(* IEC 61131-3 sources: beedance/reference (part 3) *)

FUNCTION CAUCHY : REAL
VAR_INPUT
	X : REAL;
	T : REAL;
	U : REAL;
END_VAR
VAR
	tmp: REAL;
END_VAR

tmp := x - t;
CAUCHY := math.PI_INV * U / (U*U + tmp*tmp);

(* revision hisdtory
hm	26. oct. 2008	rev 1.0
	original version

*)
END_FUNCTION

FUNCTION CAUCHYCD : REAL
VAR_INPUT
	X : REAL;
	T : REAL;
	U : REAL;
END_VAR

CAUCHYCD := 0.5 + math.PI_INV * ATAN((X - T) / U);

(* revision hisdtory
hm	26. oct. 2008	rev 1.0
	original version

*)
END_FUNCTION

FUNCTION CEIL : INT
VAR_INPUT
	X : REAL;
END_VAR

CEIL := REAL_TO_INT(x);
IF CEIL < X THEN
	CEIL := CEIL + 1;
END_IF;

END_FUNCTION

FUNCTION CEIL2 : DINT
VAR_INPUT
	X : REAL;
END_VAR

CEIL2 := REAL_TO_DINT(X);
IF DINT_TO_REAL(CEIL2) < X THEN
	CEIL2 := CEIL2 + 1;
END_IF;

END_FUNCTION

FUNCTION CMP : BOOL
VAR_INPUT
	X,Y : REAL;
	N : INT;
END_VAR
VAR
	tmp : REAL;
END_VAR

tmp := ABS(x);
IF tmp > 0.0 THEN
	tmp := EXP10(INT_TO_REAL(FLOOR(LOG(tmp))-N+1));
ELSE
	tmp := EXP10(tmp);
END_IF;
CMP := ABS(X - Y) < tmp;

END_FUNCTION

FUNCTION COSH : REAL
VAR_INPUT
	X : REAL;
END_VAR
VAR
	t: REAL;
END_VAR

T := EXP(X);
COSH := (1.0 / T + T) * 0.5;

(* revision histroy
hm	12.1.2007	rev 1.0
	original version

hm	1.12.2007	rev 1.1
	changed code to improve performance

hm	5. jan 2008	rev 1.2
	further performance improvement

hm	10. mar. 2009	rev 1.3
	real constants updated to new systax using dot
*)
END_FUNCTION

FUNCTION COTH : REAL
VAR_INPUT
	X : REAL;
END_VAR

IF X > 20.0 THEN
	COTH :=1.0;
ELSIF X < -20.0 THEN
	COTH := -1.0;
ELSE
	COTH := 1.0 + 2.0 / (EXP(X * 2.0) - 1.0);
END_IF;

(* revision histroy
hm		12.1.2007	rev 1.0
	original version

hm	1.12.2007		rev 1.1
	changed code to improve performance

hm	8. jan 2008	rev 1.2
	further improvement in performance

hm	10. mar 2008	rev 1.3
	extended range of valid inputs to +/- INV
	changed formula for better accuracy

hm	10. mar. 2009	rev 1.4
	real constants updated to new systax using dot
*)
END_FUNCTION

FUNCTION D_TRUNC : DINT
VAR_INPUT
	X : REAL;
END_VAR

D_TRUNC := REAL_TO_DINT(X);
IF X > 0.0 THEN
	IF DINT_TO_REAL(D_TRUNC) > X THEN D_TRUNC := D_TRUNC - 1; END_IF;
ELSE
	IF DINT_TO_REAL(D_TRUNC) < X THEN D_TRUNC := D_TRUNC + 1; END_IF;
END_IF;

(* for systems that support a dint truncation this routine can be replaced by trunc() *)
END_FUNCTION

FUNCTION DEC1 : INT
VAR_INPUT
	X : INT;
	N : INT;
END_VAR

IF X = 0 THEN
	DEC1 := N - 1;
ELSE
	DEC1 := X - 1;
END_IF;

(* this is a very elegant version but 50% slower
X := (X - 1 + N) MOD N;
*)
END_FUNCTION

FUNCTION DEG : REAL
VAR_INPUT
	rad : REAL;
END_VAR

DEG := MODR(57.29577951308232 * RAD, 360.0);
END_FUNCTION

FUNCTION DIFFER : BOOL
VAR_INPUT
	in1 : REAL;
	in2 : REAL;
	X : REAL;
END_VAR

DIFFER := ABS(in1 - in2) > X;
END_FUNCTION

FUNCTION ERF : REAL
VAR_INPUT
	X : REAL;
END_VAR
VAR
	x2 : REAL;
	ax2 : REAL;
END_VAR

x2 := X*X;
ax2 := 0.147 * x2 + 1.0;
ERF := SQRT(1.0 - EXP(-X2 * ((0.27323954473516 + aX2)/(ax2)))) * SGN(x);
END_FUNCTION

FUNCTION ERFC : REAL
VAR_INPUT
	X : REAL;
END_VAR

ERFC := 1.0 - ERF(X);
END_FUNCTION

FUNCTION EVEN : BOOL
VAR_INPUT
	in : DINT;
END_VAR

EVEN := NOT in.0;
END_FUNCTION

FUNCTION EXP10 : REAL
VAR_INPUT
	X : REAL;
END_VAR

EXP10 := EXP(X * 2.30258509299405);
END_FUNCTION

FUNCTION EXPN : REAL
VAR_INPUT
	X : REAL;
	N : INT;
END_VAR
VAR
	sign: BOOL;
END_VAR
VAR
	X_work : REAL;
	N_work : INT;
END_VAR
(* IEC 61131-3 does not let a POU assign to its inputs, so the body works on copies. *)
X_work := X;
N_work := N;

sign := N_work.15;
N_work := ABS(N_work);
IF N_work.0 THEN EXPN := X_work; ELSE EXPN := 1.0; END_IF;
N_work := N_work / 2;
WHILE N_work > 0 DO
   X_work := X_work * X_work;
   IF N_work.0 THEN EXPN := EXPN * X_work; END_IF;
   N_work := N_work / 2;
END_WHILE;
IF sign THEN EXPN := 1.0 / EXPN; END_IF;
END_FUNCTION

FUNCTION FACT : DINT
VAR_INPUT
	X : INT;
END_VAR

IF X >= 0 AND X <= 12 THEN
	FACT := math.FACTS[X];
ELSE
	FACT := -1;
END_IF;

(* working code without array
IF X > 12 OR X < 0 THEN
	FACT := -1;
ELSIF X < 7 THEN
	FACT := 1;
	FOR i := 2 TO X DO
		FACT := FACT * i;
	END_FOR;
ELSE
	FACT := 5040;
	FOR i := 8 TO X DO
		FACT := FACT * i;
	END_FOR;
END_IF;
*)
END_FUNCTION

FUNCTION FIB : DINT
VAR_INPUT
	X : INT;
END_VAR
VAR
	t1, t2: DINT;
END_VAR
VAR
	X_work : INT;
END_VAR
(* IEC 61131-3 does not let a POU assign to its inputs, so the body works on copies. *)
X_work := X;

IF X_work < 0 OR X_work > 46 THEN
	FIB := -1;
ELSIF X_work < 2 THEN
	FIB := X_work;
	RETURN;
ELSE
	(* the fibonacci number is the sum of the two suceeding fibonaci numbers *)
	(* we store the numbers alternatively in t1 and t2 depending on pt *)
	t2 := 1;
	WHILE X_work > 3 DO
		X_work := X_work-2;
		t1 := t1 + t2;
		t2 := t1 + t2;
	END_WHILE;
	IF X_work > 2 THEN t1 := t1 + t2; END_IF;
	fib := t1 + t2;
END_IF;

(* alternative code for very big numbers

IF X < 31 THEN
	fib := 0.4472136 * (expn(1.618034,X) - expn(-0.618034,X));
ELSE
	fib := 0.4472133 * expn(1.618034,X);
END_IF;

*)
END_FUNCTION

FUNCTION FLOOR : INT
VAR_INPUT
	X : REAL;
END_VAR

FLOOR := REAL_TO_INT(X);
IF FLOOR > X THEN
	FLOOR := FLOOR - 1;
END_IF;
END_FUNCTION

FUNCTION FLOOR2 : DINT
VAR_INPUT
	X : REAL;
END_VAR

FLOOR2 := REAL_TO_DINT(X);
IF DINT_TO_REAL(FLOOR2) > X THEN
	FLOOR2 := FLOOR2 - 1;
END_IF;
END_FUNCTION

FUNCTION FRACT : REAL
VAR_INPUT
	x : REAL;
END_VAR

IF ABS(x) < 2.0E9 THEN
	FRACT := x - DINT_TO_REAL(D_TRUNC(x));
ELSE
	FRACT := 0.0;
END_IF;
END_FUNCTION

FUNCTION GAMMA : REAL
VAR_INPUT
	X : REAL;
END_VAR

IF x > 0.0 THEN
	GAMMA := SQRT(math.PI2 / X) * EXPT(math.E_INV * (x + 1.0 / (12.0 * x - 0.1 / X)), X);
END_IF;

(* the stirling formula is not very accurate for small values of X
IF X >=0 THEN GAMMA := SQRT(math.PI2 * X) * EXPT(X / math.E, X); END_IF;
*)
END_FUNCTION

FUNCTION GAUSS : REAL
VAR_INPUT
	X : REAL;
	U : REAL;
	SI: REAL;
END_VAR
VAR
	temp: REAL;
	si_inv: REAL;
END_VAR

temp := X - U;
si_inv := 1.0  / si;
GAUSS := EXP(Temp * Temp * si_inv * si_inv * - 0.5) * 0.39894228 * si_inv;

(* revision hisdtory
hm	6. apr. 2008	rev 1.0
	original version

hm	27. oct. 2008	rev 1.1
	optimized performance

hm	10. mar. 2009	rev 1.2
	real constants updated to new systax using dot

*)
END_FUNCTION

FUNCTION GAUSSCD : REAL
VAR_INPUT
	X : REAL;
	U : REAL;
	SI: REAL;
END_VAR

GAUSSCD := (ERF((X - U) / (SI * 1.414213562)) + 1.0) * 0.5;

(* revision hisdtory
hm	6. apr. 2008	rev 1.0
	original version

hm	10. mar. 2009	rev 1.1
	real constants updated to new systax using dot

*)
END_FUNCTION

FUNCTION GCD : INT
VAR_INPUT
	A : DINT;
	B : DINT;
END_VAR
VAR
	t: DINT;
END_VAR
VAR
	A_work : DINT;
	B_work : DINT;
END_VAR
(* IEC 61131-3 does not let a POU assign to its inputs, so the body works on copies. *)
A_work := A;
B_work := B;

IF A_work = 0 THEN
	GCD := DINT_TO_INT(ABS(B_work));
ELSIF B_work = 0 THEN
	GCD := DINT_TO_INT(ABS(A_work));
ELSE
	A_work := ABS(A_work);
	B_work := ABS(B_work);
	GCD := 1;
	WHILE NOT(A_work.0 OR B_work.0) DO
		A_work := A_work / 2;
		B_work := B_work / 2;
		GCD := GCD * 2;
	END_WHILE;
	WHILE A_work > 0 DO
		IF NOT(A_work.0) THEN A_work := A_work / 2;
		ELSIF NOT(B_work.0) THEN B_work := B_work / 2;
		ELSE
			t:= ABS(A_work-B_work) / 2;
			IF A_work < B_work THEN B_work := t; ELSE A_work := T; END_IF;
		END_IF;
	END_WHILE;
	GCD := GCD * DINT_TO_INT(B_work);
END_IF;
END_FUNCTION

FUNCTION GDF : REAL
VAR_INPUT
	X : REAL;
END_VAR

IF X = 0.0 THEN
	GDF := 0.0;
ELSIF X > 15.0 THEN
	GDF := math.PI05;
ELSIF X < -15.0 THEN
	GDF := -math.PI05;
ELSE
	GDF := ATAN(EXP(X)) * 2.0 - math.PI05;
END_IF;

END_FUNCTION

FUNCTION GOLD : REAL
VAR_INPUT
	X : REAL;
END_VAR

GOLD := (X + SQRT(X*X + 4.0)) * 0.5;

END_FUNCTION

FUNCTION HYPOT : REAL
VAR_INPUT
	X : REAL;
	Y : REAL;
END_VAR

HYPOT := SQRT(x*x + y*y);

END_FUNCTION

FUNCTION INC : INT
VAR_INPUT
	X : INT;
	D : INT;
	M : INT;
END_VAR

INC := (X + D + M + 1) MOD (M + 1);
END_FUNCTION

FUNCTION INC1 : INT
VAR_INPUT
	X : INT;
	N : INT;
END_VAR

IF X >= N - 1 THEN
	INC1 := 0;
ELSE
	INC1 := X + 1;
END_IF;
END_FUNCTION

FUNCTION INC2 : INT
VAR_INPUT
	X : INT;
	D : INT;
	L : INT;
	U : INT;
END_VAR
VAR
	tmp: INT;
END_VAR

tmp := U - L + 1;
INC2 := (X + D - L + tmp) MOD tmp + L;
END_FUNCTION

FUNCTION INV : REAL
VAR_INPUT
	X : REAL;
END_VAR

IF X <> 0.0 THEN INV := 1.0 / X; END_IF;

END_FUNCTION

// Commented out for beedance: it uses REAL_TO_DW, which is commented out.
// FUNCTION LAMBERT_W : REAL
// VAR_INPUT
// 	X : REAL;
// END_VAR
// VAR
// 	w : REAL;
// 	i : INT;
// 	we: REAL;
// 	w1e: REAL;
// 	last: DWORD;
// 	ewx: REAL;
// END_VAR
//
// (* check for valid input and return -1000 if too low *)
// IF x < -0.367879441171442 THEN
// 	LAMBERT_W := -1000.0;
// 	RETURN;
// (* return 0 if x = 0 *)
// ELSIF x = 0.0 THEN
// 	RETURN;
// (* first an estimate is calculated *)
// ELSIF x <= 500.0 THEN
// 	w := LN(x + 1.0);
// 	w := 0.665 * (1.0 + 0.0195 * w) * w + 0.04;
// ELSE
// 	w := LN(x - 4.0) - (1.0 - 1.0/LN(x)) * LN(LN(x));
// END_IF;
// (* use estimate to calculate exact result *)
// FOR i := 0 TO 5 DO
// 	ewx := EXP(w);
// 	we := w * ewx - x;
// 	w1e := (w+1.0) * ewx;
// 	last := REAL_TO_DW(w) AND 16#FFFF_FFFC;
// 	w := w - (we / (w1e - (w+2.0) * we / (2.0 * w + 2.0)));
// 	IF (REAL_TO_DW(w) AND 16#FFFF_FFFC) = last THEN EXIT; END_IF;
// END_FOR;
// LAMBERT_W := w;
//
//
// (* revision hisdtory
// hm	26. oct. 2008	rev 1.0
// 	original version
//
// hm	10. mar. 2009	rev 1.1
// 	real constants updated to new systax using dot
//
// *)
// END_FUNCTION

FUNCTION LANGEVIN : REAL
VAR_INPUT
	X : REAL;
END_VAR

IF X = 0.0 THEN
	LANGEVIN := 0.0;
ELSE
	LANGEVIN := COTH(X) - 1.0 / X;
END_IF;
END_FUNCTION

FUNCTION MAX3 : REAL
VAR_INPUT
	in1 : REAL;
	in2 : REAL;
	in3 : REAL;
END_VAR

MAX3 := MAX(MAX(IN1,IN2),IN3);
END_FUNCTION

FUNCTION MID3 : REAL
VAR_INPUT
	IN1 : REAL;
	IN2 : REAL;
	IN3 : REAL;
END_VAR
VAR
	IN1_work : REAL;
	IN2_work : REAL;
END_VAR
(* IEC 61131-3 does not let a POU assign to its inputs, so the body works on copies. *)
IN1_work := IN1;
IN2_work := IN2;

IF IN1_work > IN2_work THEN MID3 := IN1_work; IN1_work := IN2_work; IN2_work := MID3; END_IF;
IF IN2_work > IN3 THEN IN2_work := IN3; END_IF;
MID3 := SEL(IN1_work > IN2_work, IN2_work, IN1_work);

(*
hm	1.1.2007	rev 1.1
	rewrote the function for better performance

hm	18. mar. 2011	rev 1.2
	improve performance
*)
END_FUNCTION

FUNCTION MIN3 : REAL
VAR_INPUT
	in1 : REAL;
	in2 : REAL;
	in3 : REAL;
END_VAR

MIN3 := MIN(MIN(IN1,IN2),IN3);
END_FUNCTION

FUNCTION MODR : REAL
VAR_INPUT
	IN : REAL;
	DIVI : REAL;
END_VAR

IF divi = 0.0 THEN
	MODR := 0.0;
ELSE
	MODR := in - DINT_TO_REAL(FLOOR2(in / divi)) * divi;
END_IF;
END_FUNCTION

FUNCTION MUL_ADD : REAL
VAR_INPUT
	X : REAL;
	K : REAL;
	O : REAL;
END_VAR

MUL_ADD := X * K + O;
END_FUNCTION

FUNCTION NEGX : REAL
VAR_INPUT
	X : REAL;
END_VAR

NEGX := -X;

END_FUNCTION

FUNCTION RAD : REAL
VAR_INPUT
	DEG : REAL;
END_VAR

RAD := MODR(0.0174532925199433 * DEG, math.PI2);
END_FUNCTION

FUNCTION RDM : REAL
VAR_INPUT
	last : REAL;
END_VAR
VAR
	tn : DWORD;
	tc : INT;
END_VAR

tn := T_PLC_MS();
tc := BIT_COUNT(tn);
tn.31 := tn.2;
tn.30 := tn.5;
tn.29 := tn.4;
tn.28 := tn.1;
tn.27 := tn.0;
tn.26 := tn.7;
tn.25 := tn.6;
tn.24 := tn.3;
tn := ROL(tn,BIT_COUNT(tn)) OR 16#80000001;
tn := ULINT_TO_DWORD(DWORD_TO_ULINT(tn) MOD 71474513 + INT_TO_ULINT(tc + 77));
RDM := FRACT(DWORD_TO_REAL(tn) / 10000000.0 * (math.E - LIMIT(0.0,last,1.0)));

(*
pt := ADR(temp);
pt^ := (T_PLC_MS() AND 16#007FFFFF) OR 16#3D000000;
RDM := fract(modR(temp*e+pi1, PI1-last) + modR(temp*PI1+e + last,e-last));
*)
END_FUNCTION

FUNCTION RDM2 : INT
VAR_INPUT
	last : INT;
	low : INT;
	high : INT;
END_VAR

RDM2 := TRUNC(RDM(FRACT(last * math.PI)) * (high - low + 1)) + low;
END_FUNCTION

FUNCTION RDMDW : DWORD
VAR_INPUT
	last : DWORD;
END_VAR
VAR
	RX: REAL;
	M: REAL;
END_VAR

M := BIT_COUNT(last);
RX := RDM(FRACT(M * math.PI));
RDMDW := SHL(REAL_TO_DWORD(rx*65535),16);
RX := RDM(FRACT(M * math.E));
RDMDW := RDMDW OR (REAL_TO_DWORD(rx*65535) AND 16#0000FFFF);
END_FUNCTION

FUNCTION REAL_TO_FRAC : FRACTION
VAR_INPUT
	X : REAL;					(* in einen Bruch umzuwandelnder Wert *)
	N : INT;					(* maximale Größe des Nenners *)
END_VAR
VAR
	temp : DINT;				(* Merker für Berechnungen *)

	sign: BOOL;					(* Vorzeichen vom Eingangswert *)
	X_gerundet: DINT;			(* Wert von Bruch, auf ganze Zahl gerundet *)
	X_ohne_Nachkomma: REAL;		(* Wert von Bruch, ohne Nachkommastellen *)
	Numerator:       DINT := 1;	(* Initialwert Zaehler  *)
	Denominator:     DINT := 0;	(* Initialwert Nenner *)
	Numerator_old:   DINT := 0;	(* Initialwert Zaehler der letzten Berechnung  *)
	Denominator_old: DINT := 1;	(* Initialwert Zaehler der letzten Berechnung   *)

END_VAR
VAR
	X_work : REAL;
END_VAR
(* IEC 61131-3 does not let a POU assign to its inputs, so the body works on copies. *)
X_work := X;

IF X_work < 0.0 THEN
	sign := TRUE;								(* Vorzeichen merken *)
	X_work := ABS(X_work);								(* Absolutwert berechnen *)
END_IF;

REPEAT
	X_gerundet := REAL_TO_DINT(X_work);

	(* Zaehler berechnen *)
	temp := numerator * X_gerundet + numerator_old;		(* Zaehler um Vorkammawert erweitern *)
	numerator_old := numerator;							(* Zaehler der letzten Berechnung speichern *)
	numerator := temp;									(* Zaehler dieser Berechnung speichern *)

	(* Nenner berechnen *)
	temp := denominator * X_gerundet + denominator_old;	(* Nenner um Vorkammawert erweitern *)
	denominator_old := denominator;						(* Nenner der letzten Berechnung speichern *)
	denominator := temp;								(* Nenner dieser Berechnung speichern *)

	(* Restwert berechnen *)
	X_ohne_Nachkomma := DINT_TO_REAL(X_gerundet);
	IF X_work = X_ohne_Nachkomma THEN						(* Bruch geht ohne Rest auf *)
		IF ABS(denominator) <= N THEN						(* kein Rundungsfehler *)
			numerator_old := numerator;					(* Numerator_old wird von Funktion zurückgegeben *)
			denominator_old := denominator;			(* Denominator_old wird von Funktion zurückgegeben *)
		END_IF
		EXIT;											(* keine weitere Berechnung notwendig *)
	ELSE
		X_work := 1.0 / (X_work - X_ohne_Nachkomma);				(* Kehrwert vom Rest -> Neuer Bruch *)
	END_IF

UNTIL
	ABS(Denominator) > N
END_REPEAT

(* correct sign if X was negative *)
IF sign THEN
	REAL_TO_FRAC.NUMERATOR := -1 * ABS(DINT_TO_INT(numerator_old));
ELSE
	REAL_TO_FRAC.NUMERATOR :=  ABS(DINT_TO_INT(numerator_old));
END_IF
REAL_TO_FRAC.DENOMINATOR := ABS(DINT_TO_INT(denominator_old));
END_FUNCTION

FUNCTION RND : REAL
VAR_INPUT
	X : REAL;
	N : INT;
END_VAR
VAR
	M : REAL;
END_VAR

IF X = 0.0 THEN
	RND := 0.0;
ELSE
	M := EXPN(10.0,N - CEIL(LOG(ABS(X))));
	RND := DINT_TO_REAL(REAL_TO_DINT(X * M)) / M;
END_IF;

END_FUNCTION

 FUNCTION ROUND : REAL
VAR_INPUT
	in : REAL;
	N : INT;
END_VAR
VAR
	X: REAL;
END_VAR

X := setup.DECADES[LIMIT(0,N,8)];
ROUND := DINT_TO_REAL(REAL_TO_DINT(in * X)) / X;

END_FUNCTION

FUNCTION SGN : INT
VAR_INPUT
	X : REAL;
END_VAR

IF X > 0 THEN
	SGN := 1;
ELSIF X < 0 THEN
	SGN := -1;
ELSE
	SGN := 0;
END_IF;

(* revision histroy
hm	16. oct 2007	rev 1.0
	original version

hm	11. nov 2007	rev 1.1
	changed type of function from real to int

*)
END_FUNCTION

FUNCTION SIGMOID : REAL
VAR_INPUT
	X : REAL;
END_VAR

IF X > 20.0 THEN
	SIGMOID := 1.0;
ELSIF x < -85.0 THEN
	SIGMOID := 0.0;
ELSE
	SIGMOID := 1.0 / (1.0 + EXP(-X));
END_IF;
END_FUNCTION

FUNCTION SIGN_I : BOOL
VAR_INPUT
	IN : DINT;
END_VAR

SIGN_I := in.31;
END_FUNCTION

FUNCTION SIGN_R : BOOL
VAR_INPUT
	in : REAL;
END_VAR

SIGN_R := in < 0.0;
END_FUNCTION

FUNCTION SINC : REAL
VAR_INPUT
	X : REAL;
END_VAR

IF X = 0.0 THEN
	SINC := 1.0;
ELSE
	SINC := SIN(x) / x;
END_IF;

(* revision histroy
hm	11. mar. 2008	rev 1.0
	original version

hm	1.12.2007	rev 1.1
	changed code to improove performance

hm 10. mar. 2009	rev 1.2
	real constants updated to new systax using dot

*)
END_FUNCTION

FUNCTION SINH : REAL
VAR_INPUT
	X : REAL;
END_VAR

IF ABS(x) < 2E-3 THEN
	SINH := X;
ELSE
	SINH := (EXP(x) - EXP(-x)) * 0.5;
END_IF;
END_FUNCTION

FUNCTION SQRTN : REAL
VAR_INPUT
	X : REAL;
	N : INT;
END_VAR

IF N > 0 THEN
	SQRTN := EXP(LN(x) / INT_TO_REAL(n));
ELSE
	SQRTN := 0.0;
END_IF;
END_FUNCTION

FUNCTION TANC : REAL
VAR_INPUT
	X : REAL;
END_VAR

IF X = 0.0 THEN
	TANC := 1.0;
ELSE
	TANC := TAN(x) / x;
END_IF;

(* revision histroy
hm	23. oct. 2008	rev 1.0
	original version

hm 10. mar. 2009	rev 1.1
	real constants updated to new systax using dot

*)
END_FUNCTION

FUNCTION TANH : REAL
VAR_INPUT
	X : REAL;
END_VAR

IF X > 20.0 THEN
	TANH := 1.0;
ELSIF X < -20.0 THEN
	TANH := -1.0;
ELSE
	TANH := 1.0 - 2.0 / (EXP(2.0 * x) + 1.0);
END_IF;

(* revision hisdtory
hm		12.1.2007		rev 1.0
	original version

hm		1.12.2007		rev 1.1
	changed code to improve performance

hm		10. mar 2008	rev 1.2
	corrected an error in formula
	extended range of valid inputs to +/- INV

hm 10. mar. 2009	rev 1.3
	real constants updated to new systax using dot

*)
END_FUNCTION

FUNCTION WINDOW : BOOL
VAR_INPUT
	low : REAL;
	in : REAL;
	high : REAL;
END_VAR

WINDOW := in < high AND in > low;
END_FUNCTION

FUNCTION WINDOW2 : BOOL
VAR_INPUT
	LOW : REAL;
	IN : REAL;
	HIGH : REAL;
END_VAR

WINDOW2 := IN >= LOW AND IN <= HIGH;
END_FUNCTION

FUNCTION_BLOCK ESR_COLLECT
VAR_INPUT
	ESR_0, ESR_1, ESR_2, ESR_3, ESR_4, ESR_5, ESR_6, ESR_7 : ARRAY [0..3] OF esr_data;
	rst : BOOL;
END_VAR
VAR_IN_OUT
	pos : INT;
END_VAR
VAR_OUTPUT
	ESR_OUT : ARRAY[0..31] OF esr_data;
END_VAR
VAR CONSTANT
	max_in : INT := 3; (* max limit of input array *)
	max_out : INT := 32; (* number of elements in array *)
END_VAR
VAR
	cnt : INT := -1;
END_VAR

IF rst OR cnt < 0 THEN
	pos := -1;
ELSE
	FOR cnt := 0 TO max_in DO
	IF esr_0[cnt].typ > 0 THEN pos := INC1(pos, max_out); esr_out[pos] := esr_0[cnt]; END_IF;
	IF esr_1[cnt].typ > 0 THEN pos := INC1(pos, max_out); esr_out[pos] := esr_1[cnt]; END_IF;
	IF esr_2[cnt].typ > 0 THEN pos := INC1(pos, max_out); esr_out[pos] := esr_2[cnt]; END_IF;
	IF esr_3[cnt].typ > 0 THEN pos := INC1(pos, max_out); esr_out[pos] := esr_3[cnt]; END_IF;
	IF esr_4[cnt].typ > 0 THEN pos := INC1(pos, max_out); esr_out[pos] := esr_4[cnt]; END_IF;
	IF esr_5[cnt].typ > 0 THEN pos := INC1(pos, max_out); esr_out[pos] := esr_5[cnt]; END_IF;
	IF esr_6[cnt].typ > 0 THEN pos := INC1(pos, max_out); esr_out[pos] := esr_6[cnt]; END_IF;
	IF esr_7[cnt].typ > 0 THEN pos := INC1(pos, max_out); esr_out[pos] := esr_7[cnt]; END_IF;
   END_FOR;
END_IF;
END_FUNCTION_BLOCK

FUNCTION_BLOCK ESR_MON_B8
VAR_INPUT
	s0, s1, s2, s3, s4, s5, s6, s7 : BOOL;
	DT_in : DT;
END_VAR
VAR_INPUT CONSTANT
	a0, a1, a2, a3, a4, a5, a6, a7 : STRING(10);
END_VAR
VAR_OUTPUT
	ESR_Flag : BOOL;
END_VAR
VAR_IN_OUT
	ESR_Out: ARRAY [0..3] OF esr_data;
END_VAR
VAR
	x0, x1, x2, x3, x4, x5, x6, x7 : BOOL;
	tx: TIME;
	cnt : INT;
END_VAR

(* read system timer *)
tx := DWORD_TO_TIME(T_PLC_MS());

ESR_Flag := FALSE;
esr_out[3].typ := 0;
esr_out[2].typ := 0;
esr_out[1].typ := 0;
esr_out[0].typ := 0;
cnt := 0;

(* check if inputs have chaged and fill buffer *)
IF s0 <> X0 THEN
	esr_out[cnt].typ := USINT_TO_BYTE(10 + BOOL_TO_USINT(s0));
	esr_out[cnt].adress := a0;
	esr_out[cnt].DS := DT_in;
	esr_out[cnt].TS := TX;
	X0 := S0;
	cnt := cnt + 1;
	esr_flag := TRUE;
END_IF;
IF s1 <> X1 THEN
	esr_out[cnt].typ := USINT_TO_BYTE(10 + BOOL_TO_USINT(s1));
	esr_out[cnt].adress := a1;
	esr_out[cnt].DS := DT_in;
	esr_out[cnt].TS := TX;
	X1 := S1;
	cnt := cnt + 1;
	esr_flag := TRUE;
END_IF;
IF s2 <> X2 THEN
	esr_out[cnt].typ := USINT_TO_BYTE(10 + BOOL_TO_USINT(s2));
	esr_out[cnt].adress := a2;
	esr_out[cnt].DS := DT_in;
	esr_out[cnt].TS := TX;
	X2 := S2;
	cnt := cnt + 1;
	esr_flag := TRUE;
END_IF;
IF s3 <> X3 THEN
	esr_out[cnt].typ := USINT_TO_BYTE(10 + BOOL_TO_USINT(s3));
	esr_out[cnt].adress := a3;
	esr_out[cnt].DS := DT_in;
	esr_out[cnt].TS := TX;
	X3 := S3;
	cnt := cnt + 1;
	esr_flag := TRUE;
END_IF;
IF s4 <> X4 AND cnt < 4 THEN
	esr_out[cnt].typ := USINT_TO_BYTE(10 + BOOL_TO_USINT(s4));
	esr_out[cnt].adress := a4;
	esr_out[cnt].DS := DT_in;
	esr_out[cnt].TS := TX;
	X4 := S4;
	cnt := cnt + 1;
	esr_flag := TRUE;
END_IF;
IF s5 <> X5  AND cnt < 4 THEN
	esr_out[cnt].typ := USINT_TO_BYTE(10 + BOOL_TO_USINT(s5));
	esr_out[cnt].adress := a5;
	esr_out[cnt].DS := DT_in;
	esr_out[cnt].TS := TX;
	X5 := S5;
	cnt := cnt + 1;
	esr_flag := TRUE;
END_IF;
IF s6 <> X6  AND cnt < 4 THEN
	esr_out[cnt].typ := USINT_TO_BYTE(10 + BOOL_TO_USINT(s6));
	esr_out[cnt].adress := a6;
	esr_out[cnt].DS := DT_in;
	esr_out[cnt].TS := TX;
	X6 := S6;
	cnt := cnt + 1;
	esr_flag := TRUE;
END_IF;
IF s7 <> X7  AND cnt < 4 THEN
	esr_out[cnt].typ := USINT_TO_BYTE(10 + BOOL_TO_USINT(s7));
	esr_out[cnt].adress := a7;
	esr_out[cnt].DS := DT_in;
	esr_out[cnt].TS := TX;
	X7 := S7;
	cnt := cnt + 1;
	esr_flag := TRUE;
END_IF;
END_FUNCTION_BLOCK

// Commented out for beedance: it reads the bits of a REAL as a DWORD, or back, through a pointer; a beedance reference (REF_TO) refers to a variable of its own type.
// FUNCTION_BLOCK ESR_MON_R4
// VAR_INPUT
// 	R0, R1, R2, R3 : REAL;
// 	DT_in : DT;
// END_VAR
// VAR_INPUT CONSTANT
// 	a0, a1, a2, a3 : STRING(10);
// 	s0, s1, s2, s3 : REAL;
// END_VAR
// VAR_OUTPUT
// 	ESR_Flag : BOOL;
// END_VAR
// VAR_IN_OUT
// 	ESR_Out: ARRAY [0..3] OF esr_data;
// END_VAR
// VAR
// 	p0, p1, p2, p3 : REF_TO DWORD;
// 	x0, x1, x2, x3 : REAL;
// 	tx: TIME;
// 	cnt : INT;
// END_VAR
//
//
// (* read system timer *)
// tx := DWORD_TO_TIME(T_PLC_MS());
// P0 := REF(R0);
// P1 := REF(R1);
// P2 := REF(R2);
// P3 := REF(R3);
//
// ESR_Flag := FALSE;
// esr_out[3].typ := 0;
// esr_out[2].typ := 0;
// esr_out[1].typ := 0;
// esr_out[0].typ := 0;
// cnt := 0;
//
// (* check if inputs have chaged and fill buffer *)
// IF DIFFER(R0,  X0, S0) THEN
// 	esr_out[cnt].typ := 20;
// 	esr_out[cnt].adress := a0;
// 	esr_out[cnt].DS := DT_in;
// 	esr_out[cnt].TS := TX;
// 	esr_out[cnt].data[0] := Byte_of_Dword(P0^,0);
// 	esr_out[cnt].data[1] := Byte_of_Dword(P0^,1);
// 	esr_out[cnt].data[2] := Byte_of_Dword(P0^,2);
// 	esr_out[cnt].data[3] := Byte_of_Dword(P0^,3);
// 	X0 := R0;
// 	cnt := cnt + 1;
// 	esr_flag := TRUE;
// END_IF;
// IF differ(R1,  X1, S1) THEN
// 	esr_out[cnt].typ := 20;
// 	esr_out[cnt].adress := a1;
// 	esr_out[cnt].DS := DT_in;
// 	esr_out[cnt].TS := TX;
// 	esr_out[cnt].data[0] := Byte_of_Dword(P1^,0);
// 	esr_out[cnt].data[1] := Byte_of_Dword(P1^,1);
// 	esr_out[cnt].data[2] := Byte_of_Dword(P1^,2);
// 	esr_out[cnt].data[3] := Byte_of_Dword(P1^,3);
// 	X1 := R1;
// 	cnt := cnt + 1;
// 	esr_flag := TRUE;
// END_IF;
// IF differ(R2,  X2, S2) THEN
// 	esr_out[cnt].typ := 20;
// 	esr_out[cnt].adress := a2;
// 	esr_out[cnt].DS := DT_in;
// 	esr_out[cnt].TS := TX;
// 	esr_out[cnt].data[0] := Byte_of_Dword(P2^,0);
// 	esr_out[cnt].data[1] := Byte_of_Dword(P2^,1);
// 	esr_out[cnt].data[2] := Byte_of_Dword(P2^,2);
// 	esr_out[cnt].data[3] := Byte_of_Dword(P2^,3);
// 	X2 := R2;
// 	cnt := cnt + 1;
// 	esr_flag := TRUE;
// END_IF;
// IF DIFFER(R3,  X3, S3) THEN
// 	esr_out[cnt].typ := 20;
// 	esr_out[cnt].adress := a3;
// 	esr_out[cnt].DS := DT_in;
// 	esr_out[cnt].TS := TX;
// 	esr_out[cnt].data[0] := Byte_of_Dword(P3^,0);
// 	esr_out[cnt].data[1] := Byte_of_Dword(P3^,1);
// 	esr_out[cnt].data[2] := Byte_of_Dword(P3^,2);
// 	esr_out[cnt].data[3] := Byte_of_Dword(P3^,3);
// 	X3 := R3;
// 	cnt := cnt + 1;
// 	esr_flag := TRUE;
// END_IF;
//
// END_FUNCTION_BLOCK

FUNCTION_BLOCK ESR_MON_X8
VAR_INPUT
	s0, s1, s2, s3, s4, s5, s6, s7 : BYTE;
	DT_in : DT;
	Mode : BYTE := 3;
END_VAR
VAR_INPUT CONSTANT
	a0, a1, a2, a3, a4, a5, a6, a7 : STRING(10);
END_VAR
VAR_OUTPUT
	ESR_Flag : BOOL;
END_VAR
VAR_IN_OUT
	ESR_Out: ARRAY [0..3] OF esr_data;
END_VAR
VAR
	x0, x1, x2, x3, x4, x5, x6, x7 : BYTE;
	tx: TIME;
	cnt : INT;
END_VAR

(* read system timer *)
tx := DWORD_TO_TIME(T_PLC_MS());

ESR_Flag := FALSE;
esr_out[3].typ := 0;
esr_out[2].typ := 0;
esr_out[1].typ := 0;
esr_out[0].typ := 0;
cnt := 0;

(* check if inputs have chaged and fill buffer *)
IF s0 <> X0 AND ((s0 < 100) OR (S0 > 99 AND S0 < 200 AND mode >= 2) OR (S0 > 199 AND mode = 3)) THEN
	esr_out[cnt] := status_to_ESR(s0, a0, DT_in, TX);
	X0 := S0;
	cnt := cnt + 1;
	esr_flag := TRUE;
END_IF;
IF s1 <> X1 AND ((s1 < 100) OR (S1 > 99 AND S1 < 200 AND mode >= 2) OR (S1 > 199 AND mode = 3)) THEN
	esr_out[cnt] := status_to_ESR(s1, a1, DT_in, TX);
	X1 := S1;
	cnt := cnt + 1;
	esr_flag := TRUE;
END_IF;
IF s2 <> X2 AND ((s2 < 100) OR (S2 > 99 AND S2 < 200 AND mode >= 2) OR (S2 > 199 AND mode = 3)) THEN
	esr_out[cnt] := status_to_ESR(s2, a2, DT_in, TX);
	X2 := S2;
	cnt := cnt + 1;
	esr_flag := TRUE;
END_IF;
IF s3 <> X3 AND ((s3 < 100) OR (S3 > 99 AND S3 < 200 AND mode >= 2) OR (S3 > 199 AND mode = 3)) THEN
	esr_out[cnt] := status_to_ESR(s3, a3, DT_in, TX);
	X3 := S3;
	cnt := cnt + 1;
	esr_flag := TRUE;
END_IF;
IF cnt < 4 AND s4 <> X4 AND ((s4 < 100) OR (S4 > 99 AND S4 < 200 AND mode >= 2) OR (S4 > 199 AND mode = 3)) THEN
	esr_out[cnt] := status_to_ESR(s4, a4, DT_in, TX);
	X4 := S4;
	cnt := cnt + 1;
	esr_flag := TRUE;
END_IF;
IF cnt < 4 AND s5 <> X5 AND ((s5 < 100) OR (S5 > 99 AND S5 < 200 AND mode >= 2) OR (S5 > 199 AND mode = 3)) THEN
	esr_out[cnt] := status_to_ESR(s5, a5, DT_in, TX);
	X5 := S5;
	cnt := cnt + 1;
	esr_flag := TRUE;
END_IF;
IF cnt < 4 AND s6 <> X6 AND ((s6 < 100) OR (S6 > 99 AND S6 < 200 AND mode >= 2) OR (S6 > 199 AND mode = 3)) THEN
	esr_out[cnt] := status_to_ESR(s6, a6, DT_in, TX);
	X6 := S6;
	cnt := cnt + 1;
	esr_flag := TRUE;
END_IF;
IF cnt < 4 AND s7 <> X7 AND ((s7 < 100) OR (S7 > 99 AND S7 < 200 AND mode >= 2) OR (S7 > 199 AND mode = 3)) THEN
	esr_out[cnt] := status_to_ESR(s7, a7, DT_in, TX);
	X7 := S7;
	cnt := cnt + 1;
	esr_flag := TRUE;
END_IF;
END_FUNCTION_BLOCK

FUNCTION OSCAT_VERSION : DWORD
VAR_INPUT
	IN : BOOL;
END_VAR

IF in THEN
	OSCAT_VERSION := DATE_TO_DWORD(D#2024-07-16);
ELSE
	OSCAT_VERSION := 335;
END_IF;
END_FUNCTION

FUNCTION STATUS_TO_ESR : esr_data
VAR_INPUT
	status : BYTE;
	adress : STRING(10);
	DT_in : DT;
	TS : TIME;
END_VAR

IF status < 100 THEN
	status_to_ESR.typ := 1;
ELSIF status < 200 THEN
	status_to_ESR.typ := 2;
ELSE
	status_to_ESR.typ := 3;
END_IF;
status_to_ESR.adress:= adress;
status_to_ESR.DS := DT_in;
status_to_ESR.TS := TS;
status_to_ESR.data[0] := status;

END_FUNCTION

// Commented out for beedance: it reads or writes the bytes of a STRING through a pointer; a beedance reference (REF_TO) refers to a whole variable of its type.
// FUNCTION BIN_TO_BYTE : BYTE
// VAR_INPUT
// 	BIN : STRING(12);
// END_VAR
// VAR
// 	pt : REF_TO BYTE;
// 	i: INT;
// 	X: BYTE;
// 	stop: INT;
// END_VAR
//
// pt := REF(bin);
// stop := LEN(bin);
// FOR I := 1 TO stop DO
// 	x := pt^;
// 	(* calculate the value of the digit *)
// 	IF X = 48 THEN
// 		BIN_TO_BYTE := SHL(BIN_TO_BYTE,1);
// 	ELSIF X = 49 THEN
// 		BIN_TO_BYTE := SHL(BIN_TO_BYTE,1) OR 1;
// 	END_IF;
// 	pt := pt + 1;
// END_FOR;
//
//
//
// (* revision histroy
// hm	18. jun. 2008	rev 1.0
// 	original release
//
// hm	20. sep. 2008	rev 1.1
// 	changed length of input string from 20 to 12
//
// hm	26. jul. 2009	rev 1.2
// 	optimized code
// *)
//
// END_FUNCTION

// Commented out for beedance: it reads or writes the bytes of a STRING through a pointer; a beedance reference (REF_TO) refers to a whole variable of its type.
// FUNCTION BIN_TO_DWORD : DWORD
// VAR_INPUT
// 	BIN : STRING(40);
// END_VAR
// VAR
// 	pt : REF_TO BYTE;
// 	i: INT;
// 	X: BYTE;
// 	stop: INT;
// END_VAR
//
// pt := REF(bin);
// stop := LEN(bin);
// FOR I := 1 TO stop DO
// 	x := pt^;
// 	(* calculate the value of the digit *)
// 	IF X = 48 THEN
// 		BIN_TO_DWORD := SHL(BIN_TO_DWORD,1);
// 	ELSIF X = 49 THEN
// 		BIN_TO_DWORD := SHL(BIN_TO_DWORD,1) OR 1;
// 	END_IF;
// 	pt := pt + 1;
// END_FOR;
//
//
//
// (* revision histroy
// hm	18. jun. 2008	rev 1.0
// 	original release
//
// hm	20. sep. 2008	rev 1.1
// 	changed length of input dtring from 20 to 40
//
// hm	26. jul 2009	rev 1.2
// 	optimized code
// *)
//
// END_FUNCTION

// Commented out for beedance: it reads or writes the bytes of a STRING through a pointer; a beedance reference (REF_TO) refers to a whole variable of its type.
// FUNCTION BYTE_TO_STRB : STRING(8)
// VAR_INPUT
// 	IN : BYTE;
// END_VAR
// VAR
// 	i: INT;
// 	pt : REF_TO BYTE;
// END_VAR
//
//
// (* pointer für die ausgabe ermitteln *)
// pt := REF(BYTE_TO_STRB);
// (* die 8 ausgabecharacter ermitteln und schreiben *)
// FOR i := 1 TO 8 DO
// 	pt^ := BOOL_TO_BYTE(in.7) + 48;
// 	in := SHL(in,1);
// 	pt := pt + 1;
// END_FOR;
//
// (* der ausgabestring muss noch mit 0 abgeschlossen werden *)
// pt^ := 0;
//
// (* code before rev 1.1
// FOR i := 1 TO 8 DO
// 	IF in.0 = 0 THEN temp := CONCAT('0', temp); ELSE temp := CONCAT('1', temp); END_IF;
// 	in := SHR(in, 1);
// END_FOR;
// BYTE_TO_STRB := temp;
// *)
// END_FUNCTION

// Commented out for beedance: it reads or writes the bytes of a STRING through a pointer; a beedance reference (REF_TO) refers to a whole variable of its type.
// FUNCTION BYTE_TO_STRH : STRING(2)
// VAR_INPUT
// 	IN : BYTE;
// END_VAR
// VAR
// 	temp : BYTE;
// 	PT : REF_TO BYTE;
// END_VAR
//
//
// (* read pointer to output string *)
// PT := REF(BYTE_TO_STRH);
// (* calculate high order hex value *)
// temp := SHR(in,4);
// (* convert value to hex character *)
// IF temp <= 9 THEN temp := temp + 48; ELSE temp := temp + 55; END_IF;
// (* write friat character to output string *)
// PT^ := temp;
// (* calculate low order hex value *)
// temp := in AND 2#00001111;
// IF temp <= 9 THEN temp := temp + 48; ELSE temp := temp + 55; END_IF;
// (* increment pointer and wirte low order character *)
// pt := pt + 1;
// pt^ := temp;
// (* set pointer at the end of the output string and close the string with 0 *)
// pt := pt + 1;
// pt^:= 0;
//
//
// (* code before rev 1.2
// FOR i := 1 TO 2 DO
// 	X := in AND 2#1111;
// 	IF X <= 9 THEN X := X + 48; ELSE X := X + 55; END_IF;
// 	Cx := CHR(X);
// 	temp := CONCAT(Cx, temp);
// 	in := SHR(in,4);
// END_FOR;
// BYTE_TO_STRH := temp;
// *)
// END_FUNCTION

// Commented out for beedance: it computes with pointers as addresses (pt := pt + 1); beedance references (REF_TO) have no arithmetic.
// FUNCTION CAPITALIZE : STRING(STRING_LENGTH)
// VAR_INPUT
// 	str : STRING(STRING_LENGTH);
// END_VAR
// VAR
// 	PT : REF_TO BYTE;
// 	pos : INT;
// 	L : INT;
// 	first : BOOL := TRUE;
// END_VAR
//
// PT := REF(CAPITALIZE);
// CAPITALIZE := str;
// L := LEN(str);
// FOR pos := 1 TO l DO
// 	IF first THEN pt^ := TO_UPPER(pt^);	END_IF;
// 	(* remember in first if the next char needs to capitalized *)
// 	first := pt^= 32;
// 	PT := pt + 1;
// END_FOR;
//
// (* revision histroy
// hm		4. mar 2008	rev 1.0
// 	original release
//
// hm	29. mar. 2008	rev 1.1
// 	changed STRING to STRING(STRING_LENGTH)
//
// hm	20. jun. 2008	rev 1.2
// 	improved performance
//
// *)
//
// END_FUNCTION

// Commented out for beedance: it uses CODE, which is commented out.
// FUNCTION CHARCODE : BYTE
// VAR_INPUT
// 	STR : STRING(10);
// END_VAR
// VAR
// 	found: STRING(1);
// 	search : STRING(10);
// 	pos: INT;
// 	i: INT;
// END_VAR
//
// IF LEN(str) = 1 THEN
// 	CHARCODE := CODE(STR, 1);
// ELSIF str <> '' THEN
// 	(* construct search string *)
// 	search := CONCAT('&', str);
// 	search := CONCAT(search, ';');
// 	WHILE pos = 0 AND (i < 4) DO
// 		i := i + 1;
// 		pos := FIND(setup.CHARNAMES[i], search);
// 	END_WHILE;
// 	found := MID(setup.CHARNAMES[i], 1, pos - 1);
// 	CHARCODE := CODE(found, 1);
// END_IF;
//
// END_FUNCTION

// Commented out for beedance: it uses CHR_TO_STRING, which is commented out.
// FUNCTION CHARNAME : STRING(10)
// VAR_INPUT
// 	C : BYTE;
// END_VAR
// VAR
// 	pos: INT;
// 	i : INT;
// END_VAR
//
// IF C <> 0 THEN
// 	(* construct search string from code followed by $ sign, also clear charname string*)
// 	CHARNAME := CHR_TO_STRING(C);
// 	CHARNAME := CONCAT(CHARNAME,'&');
// 	CHARNAME := CONCAT(';', CHARNAME);
// 	WHILE pos = 0 AND (i < 4) DO
// 		i := i + 1;
// 		pos := FIND(setup.CHARNAMES[i], CHARNAME);
// 	END_WHILE;
// 	IF pos > 0 THEN
// 		CHARNAME := MID(setup.CHARNAMES[i], 10, pos + 3);
// 		(* search for end of name and truncate *)
// 		pos := FIND(CHARNAME, ';');
// 		CHARNAME := LEFT(CHARNAME,pos - 1);
// 	ELSE
// 		CHARNAME := CHR_TO_STRING(C);
// 	END_IF;
// ELSE
// 	CHARNAME := '';
// END_IF;
//
// END_FUNCTION

// Commented out for beedance: it computes with pointers as addresses (pt := pt + 1); beedance references (REF_TO) have no arithmetic.
// FUNCTION CHR_TO_STRING : STRING(1)
// VAR_INPUT
// 	C : BYTE;
// END_VAR
// VAR
// 	PT : REF_TO BYTE;
// END_VAR
//
// PT := REF(CHR_TO_STRING);
// PT^ := C;
// pt := pt + 1;
// pt^ := 0;
// END_FUNCTION

FUNCTION CLEAN : STRING(STRING_LENGTH)
VAR_INPUT
	IN : STRING(STRING_LENGTH);
	CX : STRING(80);
END_VAR
VAR
	pos: INT := 1;
	stop: INT;
END_VAR

(* copy input string *)
CLEAN := IN;
stop := LEN(in);
WHILE pos <= stop DO
	IF FIND(cx, MID(CLEAN, 1, pos)) > 0 THEN
		(* charcter found skip to next one *)
		pos := pos + 1;
	ELSE
		(* wrong chracter needs to be deleted *)
		CLEAN := DELETE(CLEAN, 1, pos);
		stop := stop - 1;	(* the string is one character shorter now *)
	END_IF;
END_WHILE;
END_FUNCTION

// Commented out for beedance: it computes with pointers as addresses (pt := pt + 1); beedance references (REF_TO) have no arithmetic.
// FUNCTION CODE : BYTE
// VAR_INPUT
// 	STR : STRING(STRING_LENGTH);
// 	POS : INT;
// END_VAR
// VAR
// 	PT : REF_TO BYTE;
// END_VAR
//
// IF pos < 1 OR pos > LEN(str) THEN
// 	CODE := 0;
// 	RETURN;
// ELSE
// 	PT := REF(STR) + INT_TO_DWORD(pos - 1);
// 	CODE := pt^;
// END_IF;
// END_FUNCTION

// Commented out for beedance: it reads or writes the bytes of a STRING through a pointer; a beedance reference (REF_TO) refers to a whole variable of its type.
// FUNCTION COUNT_CHAR : INT
// VAR_INPUT
// 	str : STRING(STRING_LENGTH);
// 	chr : BYTE;
// END_VAR
// VAR
// 	l: INT;
// 	pt : REF_TO BYTE;
// 	pos: INT;
// END_VAR
//
// PT := REF(str);
// l := LEN(str);
// COUNT_CHAR := 0;
// FOR pos := 1 TO l DO
// 	IF pt^ = CHR THEN COUNT_CHAR := COUNT_CHAR + 1; END_IF;
//     PT := PT + 1;
// END_FOR;
// END_FUNCTION

FUNCTION COUNT_SUBSTRING : INT
VAR_INPUT
   SEARCH : STRING;
   STR : STRING;
END_VAR
VAR
   pos : INT;
   size : INT;
END_VAR
VAR
	STR_work : STRING;
END_VAR
(* IEC 61131-3 does not let a POU assign to its inputs, so the body works on copies. *)
STR_work := STR;

COUNT_SUBSTRING := 0;
size := LEN(SEARCH);
REPEAT
   pos := FIND(STR_work,SEARCH);
   IF pos > 0 THEN
      STR_work := REPLACE(STR_work, '', size,pos);
      COUNT_SUBSTRING := COUNT_SUBSTRING + 1;
   END_IF;
UNTIL pos = 0
END_REPEAT;

END_FUNCTION

// Commented out for beedance: it reads or writes the bytes of a STRING through a pointer; a beedance reference (REF_TO) refers to a whole variable of its type.
// FUNCTION DEC_TO_BYTE : BYTE
// VAR_INPUT
// 	DEC : STRING(10);
// END_VAR
// VAR
// 	pt : REF_TO BYTE;
// 	i: INT;
// 	X: BYTE;
// 	stop: INT;
// END_VAR
//
// pt := REF(dec);
// stop := LEN(DEC);
// FOR I := 1 TO stop DO
// 	(* read the first character and subtract 48 to get value in decimal 0 = 48 *)
// 	x := pt^;
// 	(* calculate the value of the digit *)
// 	IF X > 47 AND x < 58 THEN
// 		DEC_TO_BYTE := DEC_TO_BYTE * 10 + X - 48;
// 	END_IF;
// 	pt := pt + 1;
// END_FOR;
//
//
//
// (* revision histroy
// hm	20. jun. 2008	rev 1.0
// 	original release
//
// hm	30. sep.2008	rev 1.1
// 	changed length of input string from 20 to 10
// 	corrected an error where decoding of characters 8 and 9 would fail
//
// *)
//
// END_FUNCTION

// Commented out for beedance: it reads or writes the bytes of a STRING through a pointer; a beedance reference (REF_TO) refers to a whole variable of its type.
// FUNCTION DEC_TO_DWORD : DWORD
// VAR_INPUT
// 	DEC : STRING(20);
// END_VAR
// VAR
// 	pt : REF_TO BYTE;
// 	i: INT;
// 	X: BYTE;
// 	stop: INT;
// END_VAR
//
// pt := REF(dec);
// stop := LEN(dec);
// FOR I := 1 TO stop DO
// 	(* read the first character and subtract 48 to get value in decimal 0 = 48 *)
// 	x := pt^;
// 	(* calculate the value of the digit *)
// 	IF X > 47 AND x < 58 THEN
// 		DEC_TO_DWORD := DEC_TO_DWORD * 10 + X - 48;
// 	END_IF;
// 	pt := pt + 1;
// END_FOR;
//
//
//
// (* revision histroy
// hm	20. jun. 2008	rev 1.0
// 	original release
//
// hm	30. sep. 2008	rev 1.1
// 	corrected an error where decoding of characters 8 and 9 would fail
// *)
//
// END_FUNCTION

// Commented out for beedance: it reads or writes the bytes of a STRING through a pointer; a beedance reference (REF_TO) refers to a whole variable of its type.
// FUNCTION DEC_TO_INT : INT
// VAR_INPUT
// 	DEC : STRING(10);
// END_VAR
// VAR
// 	pt : REF_TO BYTE;
// 	i: INT;
// 	X: BYTE;
// 	sign: BOOL;
// 	stop: INT;
// END_VAR
//
// pt := REF(dec);
// stop := LEN(dec);
// FOR I := 1 TO stop DO
// 	(* read the first character and subtract 48 to get value in decimal 0 = 48 *)
// 	x := pt^;
// 	(* calculate the value of the digit *)
// 	IF X > 47 AND x < 58 THEN
// 		DEC_TO_INT := DEC_TO_INT * 10 + X - 48;
// 	ELSIF X = 45 AND DEC_TO_INT = 0 THEN
// 		sign := TRUE;
// 	END_IF;
// 	pt := pt + 1;
// END_FOR;
// IF sign THEN DEC_TO_INT := -DEC_TO_INT; END_IF;
//
//
// (* revision histroy
// hm	20. jun. 2008	rev 1.0
// 	original release
//
// hm	30. sep. 2008	rev 1.1
// 	changed length of input string from 20 to 10
// 	corrected an error where decoding of characters 8 and 9 would fail
// *)
//
// END_FUNCTION

FUNCTION DEL_CHARS : STRING(STRING_LENGTH)
VAR_INPUT
	IN : STRING(STRING_LENGTH);
	CX : STRING(80);
END_VAR
VAR
	pos: INT := 1;
	stop: INT;
END_VAR

(* copy input string *)
DEL_CHARS := IN;
stop := LEN(in);
WHILE pos <= stop DO
	IF FIND(cx, MID(DEL_CHARS, 1, pos)) > 0 THEN
		(* wrong chracter needs to be deleted *)
		DEL_CHARS := DELETE(DEL_CHARS, 1, pos);
		stop := stop - 1;	(* the string is one character shorter now *)
	ELSE
		(* charcter not found skip to next one *)
		pos := pos + 1;
	END_IF;
END_WHILE;
END_FUNCTION

// Commented out for beedance: it uses CODE, which is commented out.
// FUNCTION DT_TO_STRF : STRING
// VAR_INPUT
// 	DTI : DT;
// 	MS : INT;
// 	FMT : STRING;
// 	LANG : INT;
// END_VAR
// VAR CONSTANT
// 	FILL : STRING(1) := '0';
// 	BLANK : STRING(1) := ' ';
// END_VAR
// VAR
// 	ly : INT;
// 	dx: DATE;
// 	fs: STRING(10);
// 	td: TOD;
// 	tmp : INT;
// 	pos : INT;
// 	f : INT;
// END_VAR
//
// IF LANG < 1 THEN ly := language.DEFAULT; ELSE ly := MIN(language.LMAX, LANG); END_IF;
//
// (* decode date and time information *)
// dx := DT_TO_DATE(DTI);
// td := DT_TO_TOD(DTI);
//
// (* parse the format string *)
// DT_TO_STRF := FMT;
// pos := FIND(DT_TO_STRF, '#');
// WHILE pos > 0 DO
// 	(* retrieve format identifier *)
// 	f := CODE(DT_TO_STRF, pos + 1);
// 	(* generate the return string according to the format character *)
// 	fs := '';
// 	CASE f OF
// 		65 : (* letter A retunrs the year in 4 digits *)
// 			fs := INT_TO_STRING(YEAR_OF_DATE(dx));
// 		66 : (* letter B returns the year in exactly 2 digits *)
// 			fs := RIGHT(INT_TO_STRING(YEAR_OF_DATE(dx)),2);
// 		67 : (* letter C returns the month with 1 or 2 digits *)
// 			fs := INT_TO_STRING(MONTH_OF_DATE(dx));
// 		68 : (* letter D returns the month with exactly 2 digits *)
// 			fs := INT_TO_STRING(MONTH_OF_DATE(dx));
// 			IF LEN(fs) < 2 THEN fs := CONCAT('0', fs); END_IF;
// 		69 : (* letter E returns the month with 3 characters *)
// 			fs := MONTH_TO_STRING(MONTH_OF_DATE(dx), ly, 3);
// 		70 : (* letter F returns the month with all characters *)
// 			fs := MONTH_TO_STRING(MONTH_OF_DATE(dx), ly, 0);
// 		71 : (* letter G returns the day with up to 2 digits *)
// 			fs := INT_TO_STRING(DAY_OF_MONTH(dx));
// 		72 : (* letter H returns the day of the month with exactly 2 digits *)
// 			fs := INT_TO_STRING(DAY_OF_MONTH(dx));
// 			IF LEN(fs) < 2 THEN fs := CONCAT(FILL, fs); END_IF;
// 		73 : (* letter I returns the weekday as the number 1..7 1 = monday *)
// 			fs := INT_TO_STRING(DAY_OF_WEEK(dx));
// 		74 : (* letter J returns the weekday in 2 character writing *)
// 			fs := WEEKDAY_TO_STRING(DAY_OF_WEEK(dx), ly, 2);
// 		75 : (* letter K returns the weekday with all characters *)
// 			fs := WEEKDAY_TO_STRING(DAY_OF_WEEK(dx), ly, 0);
// 		76 : (* letter L returns AM or PM for the given DateTime *)
// 			IF td >= TOD#12:00:00 THEN fs := 'PM'; ELSE fs := 'AM'; END_IF;
// 		77 : (* letter M returns the hour in 1 or 2 digit form 0..24h *)
// 			fs := INT_TO_STRING(HOUR(td));
// 		78 : (* letter N returns the hour in exactly 2 digit form 0..24h *)
// 			fs := INT_TO_STRING(HOUR(td));
// 			IF LEN(fs) < 2 THEN fs := CONCAT(FILL, fs); END_IF;
// 		79 : (* letter O returns the hour in 1 or 2 digit form 0..12h *)
// 			tmp := HOUR(td) MOD 12;
// 			IF tmp = 0 THEN tmp := 12; END_IF;
// 			fs := INT_TO_STRING(tmp);
// 		80 : (* letter P returns the hour in exactly 2 digit form 0..12h *)
// 			tmp := HOUR(td) MOD 12;
// 			IF tmp = 0 THEN tmp := 12; END_IF;
// 			fs := INT_TO_STRING(tmp);
// 			IF LEN(fs) < 2 THEN fs := CONCAT(FILL, fs); END_IF;
// 		81 : (* letter Q returns the minute of the hour in 1 or two digit form *)
// 			fs := INT_TO_STRING(MINUTE(td));
// 		82 : (* letter R returns the minute of the hour in exactly two digit form *)
// 			fs := INT_TO_STRING(MINUTE(td));
// 			IF LEN(fs) < 2 THEN fs := CONCAT(FILL, fs); END_IF;
// 		83 : (* letter S returns the second of the minute in 1 or two digit form *)
// 			fs := INT_TO_STRING(REAL_TO_INT(SECOND(td)));
// 		84 : (* letter T returns the second of the minute in exactly two digit form *)
// 			fs := INT_TO_STRING(REAL_TO_INT(SECOND(td)));
// 			IF LEN(fs) < 2 THEN fs := CONCAT(FILL, fs); END_IF;
// 		85 : (* letter U returns the milliseconds in 1 to 3 digits *)
// 			fs := INT_TO_STRING(MS);
// 		86 : (* letter V returns the milliseconds in exactly 3 digit form *)
// 			fs := INT_TO_STRING(MS);
// 			fs := CONCAT('00',fs);
// 			fs := RIGHT(fs, 3);
// 		87 : (* letter W returns the day of the month with exactly 2 digits first digit is filled with blank if necessary *)
// 			fs := INT_TO_STRING(DAY_OF_MONTH(dx));
// 			IF LEN(fs) < 2 THEN fs := CONCAT(BLANK, fs); END_IF;
// 		88 : (* letter X returns the month with exactly 2 digits first digit is filled with blank if necessary *)
// 			fs := INT_TO_STRING(MONTH_OF_DATE(dx));
// 			IF LEN(fs) < 2 THEN fs := CONCAT(BLANK, fs); END_IF;
// 		END_CASE;
// 	DT_TO_STRF := REPLACE(DT_TO_STRF, fs, 2, pos);
// 	pos := FIND(DT_TO_STRF, '#');
// END_WHILE;
//
// END_FUNCTION

// Commented out for beedance: it reads or writes the bytes of a STRING through a pointer; a beedance reference (REF_TO) refers to a whole variable of its type.
// FUNCTION DWORD_TO_STRB : STRING(32)
// VAR_INPUT
// 	IN : DWORD;
// END_VAR
// VAR
// 	pt : REF_TO BYTE;
// 	i: INT;
// END_VAR
//
// (* pointer für die ausgabe ermitteln *)
// pt := REF(DWORD_TO_STRB);
// (* die 8 ausgabecharacter ermitteln und schreiben *)
// FOR i := 1 TO 32 DO
// 	pt^:= BOOL_TO_BYTE(in.31) + 48;
// 	in := SHL(in,1);
// 	pt := pt + 1;
// END_FOR;
//
// (* der ausgabestring muss nochg mit 0 abgeschlossen werden *)
// pt^ := 0;
//
// END_FUNCTION

// Commented out for beedance: it uses FIX, which is commented out.
// FUNCTION DWORD_TO_STRF : STRING(20)
// VAR_INPUT
// 	IN : DWORD;
// 	N : INT;
// END_VAR
//
//
//
// (* limit N to max 20 characters *)
// (* convert dword to string first and cut to length N *)
// DWORD_TO_STRF := FIX(DWORD_TO_STRING(in),LIMIT(0,N,20),48,1);
//
// END_FUNCTION

// Commented out for beedance: it computes with pointers as addresses (pt := pt + 1); beedance references (REF_TO) have no arithmetic.
// FUNCTION DWORD_TO_STRH : STRING(8)
// VAR_INPUT
// 	IN : DWORD;
// END_VAR
// VAR
// 	i : INT;
// 	temp : BYTE;
// 	pt : REF_TO BYTE;
// END_VAR
//
//
// (* read output adress to pointer *)
// pt := REF(DWORD_TO_STRH) + 8;
// (* wirte the closing byte for the string *)
// pt^:= 0;
//
// (* write the 8 hex characters backwards *)
// FOR i := 1 TO 8 DO;
// 	(* decrement the pointer *)
// 	pt := pt - 1;
// 	(* read the lowest order hex value *)
// 	temp := DWORD_TO_BYTE(in AND 16#0000000F);
// 	(* convert value to hex character *)
// 	IF temp <= 9 THEN temp := temp + 48; ELSE temp := temp + 55; END_IF;
// 	(* write character to output string *)
// 	PT^ := temp;
// 	(* shift in for nect hex character *)
// 	in := SHR(in,4);
// END_FOR;
//
//
// (* code beofre rev 1.2
// FOR i := 1 TO 8 DO
// 	X := DWORD_TO_BYTE(in AND 2#1111);
// 	IF X <= 9 THEN X := X + 48; ELSE X := X + 55; END_IF;
// 	Cx := CHR(X);
// 	temp := CONCAT(Cx, temp);
// 	in := SHR(in,4);
// END_FOR;
// DWORD_TO_STRH := temp;
// *)
//
// END_FUNCTION

// Commented out for beedance: it uses FINDB_NONUM, which is commented out.
// FUNCTION EXEC : STRING(STRING_LENGTH)
// VAR_INPUT
// 	str : STRING(STRING_LENGTH);
// END_VAR
// VAR
// 	pos: INT;
// 	R1: REAL;
// 	R2: REAL;
// 	operator: STRING(10);
// END_VAR
//
// (* extract both numbers and operator *)
// EXEC := UPPERCASE(TRIM(str));
//
// pos := FINDB_NONUM(EXEC);
// IF pos > 1 THEN R1 := STRING_TO_REAL(LEFT(EXEC,pos-1)); END_IF;
// R2 := STRING_TO_REAL(RIGHT(EXEC,LEN(EXEC)-pos));
// EXEC := LEFT(EXEC,pos);
// pos := FINDB_NUM(EXEC);
// operator := RIGHT(EXEC,LEN(EXEC) - pos);
// IF operator = '' AND LEN(str) = 0 THEN
// 	EXEC := '';
// 	RETURN;
// ELSIF operator = '' THEN
// 	EXEC := str;
// 	RETURN;
// END_IF;
// IF operator = '^' THEN
// 	EXEC := REAL_TO_STRING(EXPT(R1, R2));
// ELSIF operator = 'SQRT' THEN
// 	EXEC := REAL_TO_STRING(SQRT(R2));
// ELSIF operator = 'SIN' THEN
// 	EXEC := REAL_TO_STRING(SIN(r2));
// ELSIF operator = 'COS' THEN
// 	EXEC := REAL_TO_STRING(COS(r2));
// ELSIF operator = 'TAN' THEN
// 	EXEC := REAL_TO_STRING(TAN(R2));
// ELSIF operator = '*' THEN
// 	EXEC := REAL_TO_STRING(R1 * R2);
// ELSIF operator = '/' THEN
// 	IF R2 <> 0 THEN EXEC := REAL_TO_STRING(R1 / R2); ELSE EXEC := 'ERROR'; END_IF;
// ELSIF operator = '+' THEN
// 	EXEC := REAL_TO_STRING(r1 + r2);
// ELSIF operator = '-' THEN
// 	EXEC := REAL_TO_STRING(r1 - r2);
// ELSE
// 	EXEC := 'ERROR';
// END_IF;
//
// IF EXEC = 'ERROR' THEN
// 	RETURN;
// (* some systems deliver integer instead of real *)
// ELSIF FIND(EXEC,'.') = 0 THEN
// 	EXEC := CONCAT(EXEC, '.0');
// (* some systems deliver n. instead of n.0 ! *)
// ELSIF RIGHT(EXEC,1) = '.' THEN
// 	EXEC := CONCAT(EXEC,'0');
// END_IF;
// END_FUNCTION

// Commented out for beedance: it uses CHR_TO_STRING, which is commented out.
// FUNCTION FILL : STRING(STRING_LENGTH)
// VAR_INPUT
// 	C : BYTE;
// 	L : INT;
// END_VAR
// VAR
// 	i: INT;
// 	sx: STRING(1);
// END_VAR
// VAR
// 	L_work : INT;
// END_VAR
// (* IEC 61131-3 does not let a POU assign to its inputs, so the body works on copies. *)
// L_work := L;
//
// Sx := CHR_TO_STRING(c);
// (* limit L to maximum 80 characters the length of a standard string *)
// L_work := LIMIT(0,L_work,STRING_LENGTH);
// (* create a string of characters to be connected to str *)
// FOR i := 1 TO 8 DO
// 	FILL := CONCAT(FILL,FILL);
// 	IF L_work.7 THEN FILL := CONCAT(FILL,Sx); END_IF;
// 	L_work := SHL(L_work,1);
// END_FOR;
//
//
//
//
// (* revision histroy
// hm	29. mar. 2008	rev 1.0
// 	original release
//
// hm	17. dec. 2008	rev 1.1
// 	changed function chr to chr_to_string
//
// *)
// END_FUNCTION

// Commented out for beedance: it reads or writes the bytes of a STRING through a pointer; a beedance reference (REF_TO) refers to a whole variable of its type.
// FUNCTION FIND_CHAR : INT
// VAR_INPUT
// 	str : STRING(STRING_LENGTH);
// 	pos : INT;
// END_VAR
// VAR
// 	i: INT;
// 	pt : REF_TO ARRAY[1..255] OF BYTE;
// 	stop: INT;
// 	X: BYTE;
// END_VAR
//
// pt := REF(str);
// stop := LEN(str);
// FOR i := MAX(pos,1) TO stop DO;
// 	X := pt^[i];
// 	IF X > 31 AND ((setup.EXTENDED_ASCII AND X <> 127) OR (NOT setup.EXTENDED_ASCII AND X < 127)) THEN
// 		FIND_CHAR := i;
// 		RETURN;
// 	END_IF;
// END_FOR;
// FIND_CHAR := 0;
//
//
// END_FUNCTION

// Commented out for beedance: it reads or writes the bytes of a STRING through a pointer; a beedance reference (REF_TO) refers to a whole variable of its type.
// FUNCTION FIND_CTRL : INT
// VAR_INPUT
// 	str : STRING(STRING_LENGTH);
// 	pos : INT;
// END_VAR
// VAR
// 	i: INT;
// 	pt : REF_TO ARRAY[1..255] OF BYTE;
// 	stop: INT;
// 	x: BYTE;
// END_VAR
//
// pt := REF(str);
// stop := LEN(str);
// FOR i := MAX(pos,1) TO stop DO;
// 	x := PT^[I];
// 	IF x < 32 OR X = 127 THEN
// 		FIND_CTRL := i;
// 		RETURN;
// 	END_IF;
// END_FOR;
// FIND_CTRL := 0;
// END_FUNCTION

// Commented out for beedance: it reads or writes the bytes of a STRING through a pointer; a beedance reference (REF_TO) refers to a whole variable of its type.
// FUNCTION FIND_NONUM : INT
// VAR_INPUT
// 	str : STRING(STRING_LENGTH);
// 	pos : INT;
// END_VAR
// VAR
// 	i: INT;
// 	pt : REF_TO ARRAY[1..255] OF BYTE;
// 	end: INT;
// 	X: BYTE;
// END_VAR
//
// pt := REF(str);
// end := LEN(str);
// FOR i := MAX(pos,1) TO end DO;
// 	X := pt^[i];
// 	IF (X < 48 AND X <> 46) OR X > 57 THEN
// 		FIND_NONUM := i;
// 		RETURN;
// 	END_IF;
// END_FOR;
// FIND_NONUM := 0;
// END_FUNCTION

// Commented out for beedance: it reads or writes the bytes of a STRING through a pointer; a beedance reference (REF_TO) refers to a whole variable of its type.
// FUNCTION FIND_NUM : INT
// VAR_INPUT
// 	str : STRING(STRING_LENGTH);
// 	pos : INT;
// END_VAR
// VAR
// 	i : INT;
// 	pt : REF_TO ARRAY[1..255] OF BYTE;
// 	stop : INT;
// 	X: BYTE;
// END_VAR
//
// pt := REF(str);
// stop := LEN(str);
// FOR i := MAX(pos,1) TO stop DO;
// 	X := pt^[i];
// 	IF (X > 47 AND X < 58) OR X = 46 THEN
// 		FIND_NUM := i;
// 		RETURN;
// 	END_IF;
// END_FOR;
// FIND_NUM := 0;
// END_FUNCTION

FUNCTION FINDB : INT
VAR_INPUT
	str1 : STRING(STRING_LENGTH);
	str2 : STRING(STRING_LENGTH);
END_VAR
VAR
	pos: INT;
	length: INT;
END_VAR

length := LEN(str2);
FOR pos := LEN(str1) - length + 1 TO 1 BY -1 DO
	IF MID(str1,length,pos) = str2 THEN
		FindB := pos;
		RETURN;
	END_IF;
END_FOR;
FindB := 0;
END_FUNCTION

// Commented out for beedance: it computes with pointers as addresses (pt := pt + 1); beedance references (REF_TO) have no arithmetic.
// FUNCTION FINDB_NONUM : INT
// VAR_INPUT
// 	str : STRING(STRING_LENGTH);
// END_VAR
// VAR
// 	pos: INT;
// 	pt : REF_TO BYTE;
// END_VAR
//
// pt := REF(str) + LEN(str) - 1;
// FOR pos := LEN(str) TO 1 BY -1 DO;
// 	IF (PT^ < 48 AND PT^ <> 46) OR PT^ > 57 THEN
// 		FINDB_NONUM := pos;
// 		RETURN;
// 	END_IF;
// 	PT := PT - 1;
// END_FOR;
// FINDB_NONUM := 0;
// END_FUNCTION

// Commented out for beedance: it computes with pointers as addresses (pt := pt + 1); beedance references (REF_TO) have no arithmetic.
// FUNCTION FINDB_NUM : INT
// VAR_INPUT
// 	str : STRING(STRING_LENGTH);
// END_VAR
// VAR
// 	pos: INT;
// 	pt : REF_TO BYTE;
// END_VAR
//
// pt := REF(str) + LEN(str) - 1;
// FOR pos := LEN(str) TO 1 BY -1 DO;
// 	IF (PT^ > 47 AND PT^ < 58) OR PT^ = 46 THEN
// 		FINDB_NUM := pos;
// 		RETURN;
// 	END_IF;
// 	PT := PT - 1;
// END_FOR;
// FINDB_NUM := 0;
// END_FUNCTION

FUNCTION FINDP : INT
VAR_INPUT
	str : STRING(STRING_LENGTH);
	src : STRING(STRING_LENGTH);
	pos: INT;
END_VAR
VAR
	i: INT;
	ls: INT;
	lx: INT;
	stp: INT;
END_VAR

ls := LEN(str);
lx := LEN(src);
IF ls < lx OR lx = 0 THEN RETURN; END_IF;
stp := ls - lx + 1;
FOR i := MAX(pos,1) TO stp DO
	IF MID(str,lx,i) = src THEN
		FINDP := i;
		RETURN;
	END_IF;
END_FOR;
FINDP := 0;

(* revision histroy
hm	4. feb. 2008	rev 1.0
	original release

hm	29. feb 2008	rev 1.1
	ADDED MAX(pos,1) in loop initialization

hm	29. mar. 2008	rev 1.2
	changed STRING to STRING(STRING_LENGTH)
*)

END_FUNCTION

// Commented out for beedance: it uses FILL, which is commented out.
// FUNCTION FIX : STRING(STRING_LENGTH)
// VAR_INPUT
// 	str : STRING(STRING_LENGTH);
// 	L : INT;
// 	C : BYTE;
// 	M : INT;
// END_VAR
// VAR
// 	N : INT;
// 	SX: STRING(STRING_LENGTH);
// END_VAR
//
// (* make sure L does not exceed the limits of a string *)
// N := LIMIT(0,L,STRING_LENGTH) - LEN(str);
// IF N <= 0 THEN
// 	(* truncate the string at length N *)
// 	IF M = 1 THEN
// 		FIX := RIGHT(str,L);
// 	ELSE
// 		FIX := LEFT(str,L);
// 	END_IF;
// ELSIF M = 1 THEN
// 	(* connect fill characters at the beginning *)
// 	sx := FILL(C,N);
// 	FIX := CONCAT(sx,str);
// ELSIF M = 2 THEN
// 	(* center str beween fill characters *)
// 	(* for an uneven number of fill characters, there is one more at the end *)
// 	sx := FILL(C,SHR(N+1,1));
// 	FIX := CONCAT(str,sx);
// 	SX := LEFT(sx,SHR(N,1));
// 	FIX := CONCAT(sx,FIX);
// ELSE
// 	(* connect fill characters at the end *)
// 	SX := FILL(C,N);
// 	FIX := CONCAT(str,SX);
// END_IF;
//
//
// (* revision histroy
// hm	29. mar. 2008	rev 1.0
// 	original release
//
// *)
// END_FUNCTION

// Commented out for beedance: it reads or writes the bytes of a STRING through a pointer; a beedance reference (REF_TO) refers to a whole variable of its type.
// FUNCTION FLOAT_TO_REAL : REAL
// VAR_INPUT
// 	FLT : STRING(20);
// END_VAR
// VAR
// 	pt : REF_TO ARRAY[1..20] OF BYTE;
// 	i: INT;
// 	X: BYTE;
// 	sign: INT := 1;
// 	stop: INT;
// 	tmp: DINT;
// 	d : INT;
// END_VAR
//
// pt := REF(FLT);
// stop := LEN(FLT);
//
// (* we first check for sign and exit if first number or dot is reached *)
// FOR i := 1 TO stop DO
// 	X := pt^[i];
// 	IF X > 47 AND X < 58 OR X = 46 THEN
// 		EXIT;
// 	ELSIF X = 45 THEN
// 		(* code 45 is sign *)
// 		sign := -1;
// 	END_IF;
// END_FOR;
//
// (* now we scan numbers till end or dot or E is reached *)
// FOR i := i TO stop DO
// 	X := pt^[i];
// 	IF X = 44 OR X = 46 OR X = 69 OR X = 101 THEN
// 		EXIT;
// 	(* calculate the value of the digit *)
// 	ELSIF X > 47 AND x < 58 THEN
// 		tmp := tmp * 10 + X - 48;
// 	END_IF;
// END_FOR;
//
// (* process the portion after the comma if comma or dot is reached exit if exponent starts *)
// IF x = 44 OR X = 46 THEN
// 	FOR i := i + 1 TO stop DO
// 		X := pt^[i];
// 		IF X = 69 OR X = 101 THEN
// 			EXIT;
// 		ELSIF x > 47 AND x < 58 THEN
// 			tmp := tmp * 10 + X - 48;
// 			d := d - 1;
// 		END_IF;
// 	END_FOR;
// END_IF;
//
// (* process exponent if present *)
// IF X = 69 OR X = 101 THEN
// 	d := d + DEC_TO_INT(RIGHT(FLT, stop - i));
// END_IF;
//
// FLOAT_TO_REAL :=  EXPN(10, d) * DINT_TO_REAL(TMP * SIGN);
//
//
//
//
// (* revision histroy
// hm	22. jun. 2008	rev 1.0
// 	original release
//
// hm	2. oct. 2008	rev 1.1
// 	fixed an error, characters 8 and 9 would not be converted
//
// hm	22. oct. 2008	rev 1.2
// 	last fix was not done correctly
//
// hm	23. oct. 2008	rev 1.3
// 	optimzed code
// *)
//
// END_FUNCTION

// Commented out for beedance: it uses BIN_TO_BYTE, which is commented out.
// FUNCTION FSTRING_TO_BYTE : BYTE
// VAR_INPUT
// 	IN : STRING(12);
// END_VAR
//
// IF LEFT(IN, 2) = '2#' THEN
// 	(* we need to convert binary *)
// 	FSTRING_TO_BYTE := BIN_TO_BYTE(RIGHT(in, LEN(in) - 2));
// ELSIF LEFT(in, 2) = '8#' THEN
// 	(* weneed to convert octals *)
// 	FSTRING_TO_BYTE := OCT_TO_BYTE(RIGHT(in, LEN(in) - 2));
// ELSIF LEFT(in, 3) = '16#' THEN
// 	(* we need to convert hexadecimal *)
// 	FSTRING_TO_BYTE := HEX_TO_BYTE(RIGHT(in, LEN(in) - 3));
// ELSE
// 	(* we assume decimal representation *)
// 	FSTRING_TO_BYTE := DEC_TO_BYTE(CLEAN(in,'0123456789'));
// END_IF;
//
//
// (* revision histroy
// hm	18. jun. 2008	rev 1.0
// 	original release
//
// hm	20. sep. 2008	rev 1.1
// 	changed length of input string from 20 to 12
// *)
//
// END_FUNCTION

// Commented out for beedance: it uses FSTRING_TO_MONTH, which is commented out.
// FUNCTION FSTRING_TO_DT : DT
// VAR_INPUT
// 	SDT : STRING(60);
// 	FMT : STRING(60);
// END_VAR
// VAR CONSTANT
// 	ignore: STRING(1) := '*';  (* ignore character is * *)
// 	fchar : STRING(1) := '#';  (* format character is # *)
// END_VAR
// VAR
// 	c: STRING(1);
// 	tmp: STRING(20);
// 	end: INT;
// 	dy : INT := 1970;
// 	dm : INT := 1;
// 	dd : INT := 1;
// 	th : INT;
// 	tm : INT;
// 	ts : INT;
// END_VAR
// VAR
// 	SDT_work : STRING;
// 	FMT_work : STRING;
// END_VAR
// (* IEC 61131-3 does not let a POU assign to its inputs, so the body works on copies. *)
// SDT_work := SDT;
// FMT_work := FMT;
//
// (* scan input string *)
// WHILE FMT_work <> '' DO
// 	c := LEFT(FMT_work,1);
// 	IF c = ignore THEN
// 		(* skip ignore characters *)
// 		FMT_work := DELETE(FMT_work,1,1);
// 		SDT_work := DELETE(SDT_work,1,1);
// 	ELSIF C = fchar THEN
// 		(* format chracter found skip format char and read identifier *)
// 		(* store format identifier in c and skip to next char in fmt *)
// 		c := MID(FMT_work,1,2);
// 		FMT_work := DELETE(FMT_work,2,1);
// 		(* extract the substring until the end of sdt or to next char of fmt *)
// 		IF FMT_work = '' THEN
// 			tmp := SDT_work;
// 		ELSE
// 			(* serach for end of substring *)
// 			end := FIND(SDT_work, LEFT(FMT_work,1))-1;
// 			tmp := LEFT(SDT_work, end);
// 			SDT_work := DELETE(SDT_work, end,1);
// 		END_IF;
// 		(* extract information from substring *)
// 		IF c = 'Y' THEN
// 			dy := STRING_TO_INT(tmp);
// 			IF dy < 100 THEN dy := dy + 2000; END_IF;
// 		ELSIF c = 'M' THEN
// 			dm := STRING_TO_INT(tmp);
// 		ELSIF c = 'N' THEN
// 			dm := FSTRING_TO_MONTH(tmp,0);
// 		ELSIF c = 'D' THEN
// 			dd := STRING_TO_INT(tmp);
// 		ELSIF c = 'h' THEN
// 			th := STRING_TO_INT(tmp);
// 		ELSIF c = 'm' THEN
// 			tm := STRING_TO_INT(tmp);
// 		ELSIF c = 's' THEN
// 			ts := STRING_TO_INT(tmp);
// 		END_IF;
// 	ELSIF c = LEFT(SDT_work,1) THEN
// 		(* skip matching characters *)
// 		FMT_work := DELETE(FMT_work,1,1);
// 		SDT_work := DELETE(SDT_work,1,1);
// 	ELSE
// 		RETURN;
// 	END_IF;
// END_WHILE;
//
// FSTRING_TO_DT := SET_DT(dy,dm,dd,th,tm,ts);
//
//
// (* revision histroy
// hm	24. sep. 2008	rev 1.0
// 	original release
//
//
// *)
//
// END_FUNCTION

// Commented out for beedance: it uses BIN_TO_DWORD, which is commented out.
// FUNCTION FSTRING_TO_DWORD : DWORD
// VAR_INPUT
// 	IN : STRING(40);
// END_VAR
//
// IF LEFT(IN, 2) = '2#' THEN
// 	(* we need to convert binary *)
// 	FSTRING_TO_DWORD := BIN_TO_DWORD(RIGHT(in, LEN(in) - 2));
// ELSIF LEFT(in, 2) = '8#' THEN
// 	(* weneed to convert octals *)
// 	FSTRING_TO_DWORD := OCT_TO_DWORD(RIGHT(in, LEN(in) - 2));
// ELSIF LEFT(in, 3) = '16#' THEN
// 	(* we need to convert hexadecimal *)
// 	FSTRING_TO_DWORD := HEX_TO_DWORD(RIGHT(in, LEN(in) - 3));
// ELSE
// 	(* we assume decimal representation *)
// 	FSTRING_TO_DWORD := DEC_TO_DWORD(CLEAN(in,'0123456789'));
// END_IF;
//
//
// (* revision histroy
// hm	18. jun. 2008	rev 1.0
// 	original release
//
// hm	20. sep. 2008	rev 1.1
// 	changed length of input dtring from 20 to 40
//
//
// *)
//
// END_FUNCTION

// Commented out for beedance: it uses CAPITALIZE, which is commented out.
// FUNCTION FSTRING_TO_MONTH : INT
// VAR_INPUT
// 	MTH : STRING(20);
// 	LANG : INT;
// END_VAR
// VAR
// 	lx: INT;
// END_VAR
// VAR
// 	MTH_work : STRING;
// END_VAR
// (* IEC 61131-3 does not let a POU assign to its inputs, so the body works on copies. *)
// MTH_work := MTH;
//
// IF LANG = 0 THEN lx := LANGUAGE.DEFAULT; ELSE lx := MIN(LANG, LANGUAGE.LMAX); END_IF;
// MTH_work := TRIM(MTH_work);
// MTH_work := CAPITALIZE(LOWERCASE(MTH_work));
//
// FOR FSTRING_TO_MONTH := 1 TO 12 DO
// 	IF MTH_work = language.MONTHS[lx, FSTRING_TO_MONTH] THEN RETURN; END_IF;
// 	IF MTH_work = language.MONTHS3[lx, FSTRING_TO_MONTH] THEN RETURN; END_IF;
// END_FOR;
//
// (* since no name matched try to decode as integer *)
// FSTRING_TO_MONTH := STRING_TO_INT(MTH_work);
//
//
//
//
// (* revision histroy
// hm	25. sep. 2008	rev 1.0
// 	original release
//
// hm	19. oct. 2008	rev 1.1
// 	changed language setup constants
//
// hm	25. oct. 2008	rev 1.2
// 	optimized code
// *)
//
// END_FUNCTION

// Commented out for beedance: it uses FSTRING_TO_WEEKDAY, which is commented out.
// FUNCTION FSTRING_TO_WEEK : BYTE
// VAR_INPUT
// 	WEEK : STRING(60);
// 	LANG : INT;
// END_VAR
// VAR
// 	pos: INT;
// END_VAR
// VAR
// 	WEEK_work : STRING;
// END_VAR
// (* IEC 61131-3 does not let a POU assign to its inputs, so the body works on copies. *)
// WEEK_work := WEEK;
//
// pos := FIND(WEEK_work, ',');
// WHILE pos > 0 DO
// 	FSTRING_TO_WEEK := FSTRING_TO_WEEK OR SHR(BYTE#128, FSTRING_TO_WEEKDAY(MID(WEEK_work, pos - 1, 1), LANG));
// 	WEEK_work := RIGHT(WEEK_work, LEN(WEEK_work) - pos);
// 	pos := FIND(WEEK_work, ',');
// END_WHILE;
// FSTRING_TO_WEEK := (FSTRING_TO_WEEK OR SHR(BYTE#128, FSTRING_TO_WEEKDAY(WEEK_work, LANG))) AND BYTE#127;
//
//
// (* revision histroy
// hm	18. jun. 2008	rev 1.0
// 	original release
//
// hm	25. oct. 2008	rev 1.1
// 	using language defauls and input lang
// *)
//
// END_FUNCTION

// Commented out for beedance: it uses CAPITALIZE, which is commented out.
// FUNCTION FSTRING_TO_WEEKDAY : INT
// VAR_INPUT
// 	WDAY : STRING(20);
// 	LANG : INT;
// END_VAR
// VAR
// 	tmp: STRING(2);
// 	i: INT;
// 	ly: INT;
// END_VAR
//
// IF LANG = 0 THEN ly := LANGUAGE.DEFAULT; ELSE ly := MIN(LANG, LANGUAGE.LMAX); END_IF;
// (* tmp needs to be calculated first otherwise find can return wrong values *)
// tmp := TRIM(wday);
// tmp := CAPITALIZE(LOWERCASE(tmp));
// FOR i := 1 TO 7 DO
// 	IF language.WEEKDAYS2[ly, i] = tmp THEN
// 		FSTRING_TO_WEEKDAY := i;
// 		RETURN;
// 	END_IF;
// END_FOR;
// FSTRING_TO_WEEKDAY := STRING_TO_INT(WDAY);
//
//
//
//
// (* revision histroy
// hm	18. jun. 2008	rev 1.0
// 	original release
//
// hm	18. jul. 2008	rev 1.1
// 	changed nested call of left(trim()) for compatibility reasons
//
// hm	25. oct. 2008	rev 1.2
// 	using language constants
// *)
//
// END_FUNCTION

// Commented out for beedance: it reads or writes the bytes of a STRING through a pointer; a beedance reference (REF_TO) refers to a whole variable of its type.
// FUNCTION HEX_TO_BYTE : BYTE
// VAR_INPUT
// 	HEX : STRING(5);
// END_VAR
// VAR
// 	pt : REF_TO BYTE;
// 	i: INT;
// 	X: BYTE;
// 	stop: INT;
// END_VAR
//
// pt := REF(hex);
// stop := LEN(hex);
// FOR I := 1 TO stop DO
// 	(* read the first character and subtract 48 to get value in decimal 0 = 48 *)
// 	x := pt^;
// 	(* calculate the value of the digit *)
// 	IF X > 47 AND x < 58 THEN
// 		HEX_TO_BYTE := SHL(HEX_TO_BYTE,4) + X - 48;
// 	ELSIF X > 64 AND X < 71 THEN
// 		HEX_TO_BYTE := SHL(HEX_TO_BYTE,4) + X - 55;
// 	ELSIF X > 96 AND X < 103 THEN
// 		HEX_TO_BYTE := SHL(HEX_TO_BYTE,4) + X - 87;
// 	END_IF;
// 	pt := pt + 1;
// END_FOR;
//
//
//
//
// (* revision histroy
// hm	18. jun. 2008	rev 1.0
// 	original release
//
// hm	20. sep.2008	rev 1.1
// 	changed length of input string from 20 to 5
//
// *)
//
// END_FUNCTION

// Commented out for beedance: it reads or writes the bytes of a STRING through a pointer; a beedance reference (REF_TO) refers to a whole variable of its type.
// FUNCTION HEX_TO_DWORD : DWORD
// VAR_INPUT
// 	Hex : STRING(20);
// END_VAR
// VAR
// 	pt : REF_TO BYTE;
// 	i: INT;
// 	X: BYTE;
// 	stop: INT;
// END_VAR
//
// pt := REF(hex);
// stop := LEN(hex);
// FOR I := 1 TO stop DO
// 	(* read the first character and subtract 48 to get value in decimal 0 = 48 *)
// 	x := pt^;
// 	(* calculate the value of the digit *)
// 	IF X > 47 AND x < 58 THEN
// 		HEX_TO_DWORD := SHL(HEX_TO_DWORD,4) + X - 48;
// 	ELSIF X > 64 AND X < 71 THEN
// 		HEX_TO_DWORD := SHL(HEX_TO_DWORD,4) + X - 55;
// 	ELSIF X > 96 AND X < 103 THEN
// 		HEX_TO_DWORD := SHL(HEX_TO_DWORD,4) + X - 87;
// 	END_IF;
// 	pt := pt + 1;
// END_FOR;
//
//
//
// (* revision histroy
// hm	2.10.2007		rev 1.0
// 	original release
//
// hm	19.11.2007		rev 1.1
// 	changed type of function from int to dword
//
// hm 	4. mar 2008		rev 1.2
// 	added support for a..f and return 0 for invalid string
//
// hm	29. mar. 2008	rev 1.3
// 	changed STRING to STRING(8)
//
// hm	18. jun. 2008	rev 1.4
// 	changed input hex to STRING(20)
// 	function now ignores wrong characters
// *)
//
// END_FUNCTION

// Commented out for beedance: it reads or writes the bytes of a STRING through a pointer; a beedance reference (REF_TO) refers to a whole variable of its type.
// FUNCTION IS_ALNUM : BOOL
// VAR_INPUT
// 	str : STRING(STRING_LENGTH);
// END_VAR
// VAR
// 	L: INT;
// 	pt : REF_TO BYTE;
// 	pos: INT;
// END_VAR
//
// PT := REF(str);
// L := LEN(str);
// FOR pos := 1 TO L DO
// 	IF NOT (ISC_ALPHA(pt^) OR ISC_NUM(pt^)) THEN
// 		IS_ALNUM := FALSE;
// 		RETURN;
// 	END_IF;
//     	PT := PT + 1;
// END_FOR;
// IS_ALNUM := L > 0;
// END_FUNCTION

// Commented out for beedance: it reads or writes the bytes of a STRING through a pointer; a beedance reference (REF_TO) refers to a whole variable of its type.
// FUNCTION IS_ALPHA : BOOL
// VAR_INPUT
// 	str : STRING(STRING_LENGTH);
// END_VAR
// VAR
// 	L: INT;
// 	pt : REF_TO BYTE;
// 	pos: INT;
// END_VAR
//
// PT := REF(str);
// L := LEN(str);
// FOR pos := 1 TO L DO
// 	IF NOT ISC_ALPHA(pt^) THEN
// 		IS_ALPHA := FALSE;
// 		RETURN;
// 	END_IF;
//     	PT := PT + 1;
// END_FOR;
// IS_ALPHA := L > 0;
// END_FUNCTION

FUNCTION IS_CC : BOOL
VAR_INPUT
	str : STRING(STRING_LENGTH);
	cmp : STRING(STRING_LENGTH);
END_VAR
VAR
	L: INT;
	pos: INT;
END_VAR

L := LEN(str);
FOR pos := 1 TO L DO
	IF FIND(CMP,MID(str,1,pos)) = 0 THEN RETURN; END_IF;
END_FOR;
IS_CC := L > 0;
END_FUNCTION

// Commented out for beedance: it reads or writes the bytes of a STRING through a pointer; a beedance reference (REF_TO) refers to a whole variable of its type.
// FUNCTION IS_CTRL : BOOL
// VAR_INPUT
// 	STR : STRING(STRING_LENGTH);
// END_VAR
// VAR
// 	L: INT;
// 	pt : REF_TO BYTE;
// 	pos: INT;
// END_VAR
//
// PT := REF(str);
// L := LEN(str);
// FOR pos := 1 TO L DO
// 	IF NOT (ISC_CTRL(pt^)) THEN
// 		IS_CTRL := FALSE;
// 		RETURN;
// 	END_IF;
//     	PT := PT + 1;
// END_FOR;
// IS_CTRL := L > 0;
// END_FUNCTION

// Commented out for beedance: it reads or writes the bytes of a STRING through a pointer; a beedance reference (REF_TO) refers to a whole variable of its type.
// FUNCTION IS_HEX : BOOL
// VAR_INPUT
// 	str : STRING(STRING_LENGTH);
// END_VAR
// VAR
// 	L: INT;
// 	pt : REF_TO BYTE;
// 	pos: INT;
// END_VAR
//
// PT := REF(str);
// L := LEN(str);
// FOR pos := 1 TO L DO
// 	IF NOT (ISC_HEX(pt^)) THEN
// 		IS_HEX := FALSE;
// 		RETURN;
// 	END_IF;
//     	PT := PT + 1;
// END_FOR;
// IS_HEX := L > 0;
// END_FUNCTION

// Commented out for beedance: it reads or writes the bytes of a STRING through a pointer; a beedance reference (REF_TO) refers to a whole variable of its type.
// FUNCTION IS_LOWER : BOOL
// VAR_INPUT
// 	str : STRING(STRING_LENGTH);
// END_VAR
// VAR
// 	l: INT;
// 	pt : REF_TO BYTE;
// 	pos: INT;
// END_VAR
//
// PT := REF(str);
// L := LEN(str);
// FOR pos := 1 TO L DO
// 	IF NOT (ISC_LOWER(pt^)) THEN
// 		IS_LOWER := FALSE;
// 		RETURN;
// 	END_IF;
//     	PT := PT + 1;
// END_FOR;
// IS_LOWER := L > 0;
// END_FUNCTION

FUNCTION IS_NCC : BOOL
VAR_INPUT
	str : STRING(STRING_LENGTH);
	cmp : STRING(STRING_LENGTH);
END_VAR
VAR
	L: INT;
	pos: INT;
END_VAR

L := LEN(str);
FOR pos := 1 TO L DO
	IF FIND(CMP,MID(str,1,pos)) > 0 THEN RETURN; END_IF;
END_FOR;
IS_NCC := TRUE;
END_FUNCTION

// Commented out for beedance: it reads or writes the bytes of a STRING through a pointer; a beedance reference (REF_TO) refers to a whole variable of its type.
// FUNCTION IS_NUM : BOOL
// VAR_INPUT
// 	str : STRING(STRING_LENGTH);
// END_VAR
// VAR
// 	L : INT;
// 	pt : REF_TO BYTE;
// 	pos: INT;
// END_VAR
//
// PT := REF(str);
// L := LEN(str);
// FOR pos := 1 TO L DO
// 	IF NOT (ISC_NUM(pt^)) THEN
// 		IS_NUM := FALSE;
// 		RETURN;
// 	END_IF;
//     	PT := PT + 1;
// END_FOR;
// IS_NUM := L > 0;
// END_FUNCTION

// Commented out for beedance: it reads or writes the bytes of a STRING through a pointer; a beedance reference (REF_TO) refers to a whole variable of its type.
// FUNCTION IS_UPPER : BOOL
// VAR_INPUT
// 	str : STRING(STRING_LENGTH);
// END_VAR
// VAR
// 	L: INT;
// 	pt : REF_TO BYTE;
// 	pos: INT;
// END_VAR
//
// PT := REF(str);
// L := LEN(str);
// FOR pos := 1 TO L DO
// 	IF NOT (ISC_UPPER(pt^)) THEN
// 		IS_UPPER := FALSE;
// 		RETURN;
// 	END_IF;
//     	PT := PT + 1;
// END_FOR;
// IS_UPPER := L > 0;
// END_FUNCTION

FUNCTION ISC_ALPHA : BOOL
VAR_INPUT
	IN : BYTE;
END_VAR

IF setup.EXTENDED_ASCII THEN
	ISC_ALPHA := (in > 64 AND in < 91) OR (in > 191  AND in <> 215 AND in <> 247) OR (in > 96 AND in < 123);
ELSE
	ISC_ALPHA := (IN > 64 AND IN < 91) OR (in > 96 AND in < 123);
END_IF;

END_FUNCTION

FUNCTION ISC_CTRL : BOOL
VAR_INPUT
	IN : BYTE;
END_VAR

ISC_CTRL := IN < 32 OR IN = 127;
END_FUNCTION

FUNCTION ISC_HEX : BOOL
VAR_INPUT
	IN : BYTE;
END_VAR

ISC_HEX := (IN > 47 AND IN < 58) OR (IN > 64 AND IN < 71) OR (IN > 96 AND IN < 103);
END_FUNCTION

FUNCTION ISC_LOWER : BOOL
VAR_INPUT
	IN : BYTE;
END_VAR

IF setup.EXTENDED_ASCII THEN
	ISC_LOWER := ((in > 96) AND (in < 123)) OR ((in > 222) AND (in <> 247));
ELSE
	ISC_LOWER := ((in > 96) AND (in < 123));
END_IF;
END_FUNCTION

FUNCTION ISC_NUM : BOOL
VAR_INPUT
	IN : BYTE;
END_VAR

ISC_NUM := IN > 47 AND IN < 58;
END_FUNCTION

FUNCTION ISC_UPPER : BOOL
VAR_INPUT
	IN : BYTE;
END_VAR

IF setup.EXTENDED_ASCII THEN
	ISC_UPPER :=  ((in > 64) AND (in < 91)) OR (((in > 191) AND (in < 223)) AND (in <> 215));
ELSE
	ISC_UPPER := ((in > 64) AND (in < 91));
END_IF;
END_FUNCTION

// Commented out for beedance: it computes with pointers as addresses (pt := pt + 1); beedance references (REF_TO) have no arithmetic.
// FUNCTION LOWERCASE : STRING(STRING_LENGTH)
// VAR_INPUT
// 	str : STRING(STRING_LENGTH);
// END_VAR
// VAR
// 	PT : REF_TO BYTE;
// 	pos: INT;
// 	l: INT;
// END_VAR
//
// PT := REF(LOWERCASE);
// lowercase := str;
// l := LEN(str);
// FOR pos := 1 TO l DO
// 	pt^ := TO_LOWER(pt^);
// 	PT := PT + 1;
// END_FOR;
//
// (* revision histroy
// hm	6. oct. 2006	rev 1.0
// 	original release
//
// hm	4. feb. 2008	rev 1.1
// 	improved performance
// 	added Ä.Ö,Ü
//
// hm	6. mar. 2008	rev 1.2
// 	added support for exteded Ascii
//
// hm	29. mar. 2008	rev 1.3
// 	changed STRING to STRING(STRING_LENGTH)
// *)
//
// END_FUNCTION

FUNCTION_BLOCK MESSAGE_4R
VAR_INPUT
	M0 : STRING(STRING_LENGTH);
	M1 : STRING(STRING_LENGTH);
	M2 : STRING(STRING_LENGTH);
	M3 : STRING(STRING_LENGTH);
	MM : INT := 3;
	ENQ : BOOL := TRUE;
	CLK : BOOL := TRUE;
	T1 : TIME := T#3s;
END_VAR
VAR_OUTPUT
	MX : STRING(STRING_LENGTH);
	MN : INT;
	TR : BOOL;
END_VAR
VAR
	timer : TON;
	edge: BOOL;
END_VAR

(* check for rising edge on EN *)
TR := FALSE;
IF ENQ THEN
	IF (NOT edge AND clk) OR timer.q THEN
			MN := INC1(MN, MM);
			TR := TRUE;
			timer(in := FALSE);
			CASE MN OF
				0 : MX := M0;
				1 : MX := M1;
				2 : MX := M2;
				3 : MX := M3;
			END_CASE;
	END_IF;
	edge := clk;
	timer( in := CLK, pt := T1);
ELSE
	MX := '';
	MN := 0;
END_IF;

END_FUNCTION_BLOCK

FUNCTION_BLOCK MESSAGE_8
VAR_INPUT
	IN1 : BOOL;
	IN2 : BOOL;
	IN3 : BOOL;
	IN4 : BOOL;
	IN5 : BOOL;
	IN6 : BOOL;
	IN7 : BOOL;
	IN8 : BOOL;
END_VAR
VAR_INPUT CONSTANT
	S1 : STRING(STRING_LENGTH);
	S2 : STRING(STRING_LENGTH);
	S3 : STRING(STRING_LENGTH);
	S4 : STRING(STRING_LENGTH);
	S5 : STRING(STRING_LENGTH);
	S6 : STRING(STRING_LENGTH);
	S7 : STRING(STRING_LENGTH);
	S8 : STRING(STRING_LENGTH);
END_VAR
VAR_OUTPUT
	M : STRING(STRING_LENGTH);
END_VAR

(* check if an alarm is present if yes set the output M otherwise clear M *)
IF in1 THEN
	M := S1;
ELSIF in2 THEN
	M := S2;
ELSIF in3 THEN
	M := S3;
ELSIF in4 THEN
	M := S4;
ELSIF in5 THEN
	M := S5;
ELSIF in6 THEN
	M := S6;
ELSIF in7 THEN
	M := S7;
ELSIF in8 THEN
	M := S8;
ELSE
	M := '';
END_IF;

END_FUNCTION_BLOCK

// Commented out for beedance: it reads or writes the bytes of a STRING through a pointer; a beedance reference (REF_TO) refers to a whole variable of its type.
// FUNCTION MIRROR : STRING(STRING_LENGTH)
// VAR_INPUT
// 	str : STRING(STRING_LENGTH);
// END_VAR
// VAR
// 	pi : REF_TO ARRAY[1..255] OF BYTE;
// 	po : REF_TO BYTE;
// 	lx: INT;
// 	i: INT;
// END_VAR
//
// pi := REF(str);
// po := REF(mirror);
// lx := LEN(str);
// FOR i := lx TO 1 BY - 1 DO
// 	po^ := pi^[i];
// 	po := po + 1;
// END_FOR;
// (* close output string *)
// po^:= 0;
//
//
// (* revision histroy
// hm	4. feb. 2008	rev 1.0
// 	original release
//
// hm	29. mar. 2008	rev 1.1
// 	changed STRING to STRING(STRING_LENGTH)
// *)
//
// END_FUNCTION

FUNCTION MONTH_TO_STRING : STRING(10)
VAR_INPUT
	MTH : INT;
	LANG : INT;
	LX : INT;
END_VAR
VAR
	ly : INT;
END_VAR

IF LANG <= 0 THEN Ly := LANGUAGE.DEFAULT; ELSE ly := MIN(LANG, language.LMAX); END_IF;
IF MTH < 1 OR MTH > 12 THEN
	RETURN;
ELSIF LX = 0 THEN
	MONTH_TO_STRING := language.MONTHS[ly, MTH];
ELSIF Lx = 3 THEN
	MONTH_TO_STRING := language.MONTHS3[ly, MTH];
END_IF;

(* revisison history

hm	21. sep. 2008	rev 1.0
	original version

hm	19. oct. 2008	rev 1.1
	changed language setup constants

hm 16.  jul 2024   rev 1.2
       addaed boundary check to respect array limits
*)
END_FUNCTION

// Commented out for beedance: it reads or writes the bytes of a STRING through a pointer; a beedance reference (REF_TO) refers to a whole variable of its type.
// FUNCTION OCT_TO_BYTE : BYTE
// VAR_INPUT
// 	OCT : STRING(10);
// END_VAR
// VAR
// 	pt : REF_TO BYTE;
// 	i: INT;
// 	X: BYTE;
// 	stop: INT;
// END_VAR
//
// pt := REF(oct);
// stop := LEN(oct);
// FOR I := 1 TO stop DO
// 	(* read the first character and subtract 48 to get value in decimal 0 = 48 *)
// 	x := pt^;
// 	(* calculate the value of the digit *)
// 	IF X > 47 AND x < 56 THEN
// 		OCT_TO_BYTE := SHL(OCT_TO_BYTE,3) + X - 48;
// 	END_IF;
// 	pt := pt + 1;
// END_FOR;
//
//
//
// (* revision histroy
// hm	18. jun. 2008	rev 1.0
// 	original release
//
// hm	20. sep. 2008	rev 1.1
// 	changed length of input string from 20 to 10
//
// *)
//
// END_FUNCTION

// Commented out for beedance: it reads or writes the bytes of a STRING through a pointer; a beedance reference (REF_TO) refers to a whole variable of its type.
// FUNCTION OCT_TO_DWORD : DWORD
// VAR_INPUT
// 	OCT : STRING(20);
// END_VAR
// VAR
// 	pt : REF_TO BYTE;
// 	i: INT;
// 	X: BYTE;
// 	stop: INT;
// END_VAR
//
// pt := REF(oct);
// stop := LEN(oct);
// FOR I := 1 TO stop DO
// 	(* read the first character and subtract 48 to get value in decimal 0 = 48 *)
// 	x := pt^;
// 	(* calculate the value of the digit *)
// 	IF X > 47 AND x < 56 THEN
// 		OCT_TO_DWORD := SHL(OCT_TO_DWORD,3) + X - 48;
// 	END_IF;
// 	pt := pt + 1;
// END_FOR;
//
//
//
//
// (* revision histroy
// hm	18. jun. 2008	rev 1.0
// 	original release
//
//
// *)
//
// END_FUNCTION

FUNCTION REAL_TO_STRF : STRING(20)
VAR_INPUT
	IN : REAL;
	N : INT;
	D : STRING(1);
END_VAR
VAR
	O: REAL;
	i: INT;
END_VAR
VAR
	N_work : INT;
END_VAR
(* IEC 61131-3 does not let a POU assign to its inputs, so the body works on copies. *)
N_work := N;

(* LIMIT N to 0 .. 7 *)
N_work := LIMIT(0,N_work,7);
(* round the input to N digits and convert to string *)
O := ABS(in) * EXP10(N_work);
REAL_TO_STRF := DINT_TO_STRING(REAL_TO_DINT(O));
(* add zeroes in front to make sure sting is at least 8 digits long *)
FOR i := LEN(REAL_TO_STRF) TO N_work DO REAL_TO_STRF := CONCAT('0', REAL_TO_STRF); END_FOR;
(* add a dot if n > 0 *)
IF N_work > 0 THEN REAL_TO_STRF := INSERT(REAL_TO_STRF, D, LEN(REAL_TO_STRF) - N_work); END_IF;
(* add a minus sign if in is negative *)
IF in < 0 THEN REAL_TO_STRF := CONCAT('-', REAL_TO_STRF); END_IF;

END_FUNCTION

FUNCTION REPLACE_ALL : STRING(STRING_LENGTH)
VAR_INPUT
	str : STRING(STRING_LENGTH);
	src : STRING(STRING_LENGTH);
	rep : STRING(STRING_LENGTH);
END_VAR
VAR
	pos: INT;
	lp : INT;
	lx : INT;
END_VAR

REPLACE_ALL := str;
lx := LEN(src);
lp := LEN(rep);
pos := FINDP(REPLACE_ALL, src, 1);
WHILE pos > 0 DO
	REPLACE_ALL := REPLACE(REPLACE_ALL,rep,lx, pos);
	pos := FINDP(REPLACE_ALL, src, pos + lp);
END_WHILE;

(* revision histroy
hm	4. feb. 2008	rev 1.0
	original release

hm	29. mar. 2008	rev 1.1
	changed STRING to STRING(STRING_LENGTH)
*)

END_FUNCTION

FUNCTION REPLACE_CHARS : STRING(STRING_LENGTH)
VAR_INPUT
	STR : STRING(STRING_LENGTH);
	SRC : STRING;
	REP : STRING;
END_VAR
VAR
	a, b : INT;
	c: STRING(1);
	stp: INT;
END_VAR
VAR
	SRC_work : STRING;
	REP_work : STRING;
END_VAR
(* IEC 61131-3 does not let a POU assign to its inputs, so the body works on copies. *)
SRC_work := SRC;
REP_work := REP;

REPLACE_CHARS := STR;
(* make sure rep and src are of same length and length is > 0 *)
a := LEN(SRC_work);
b := LEN(REP_work);
IF a < b THEN
	REP_work := LEFT(REP_work, a);
ELSIF b < a THEN
	SRC_work := LEFT(SRC_work, b);
END_IF;

(* search the string and replace if necessary *)
stp := LEN(str);
FOR a := 1 TO stp DO
	c := MID(REPLACE_CHARS, 1, a);
	b := FIND(SRC_work, c);
	IF b > 0 THEN
		REPLACE_CHARS := REPLACE(REPLACE_CHARS, MID(REP_work, 1, b), 1, a);
	END_IF;
END_FOR;

END_FUNCTION

// Commented out for beedance: it reads or writes the bytes of a STRING through a pointer; a beedance reference (REF_TO) refers to a whole variable of its type.
// FUNCTION REPLACE_UML : STRING(STRING_LENGTH)
// VAR_INPUT
// 	str : STRING(STRING_LENGTH);
// END_VAR
// VAR
// 	L : INT;
// 	pt : REF_TO BYTE;
// 	pto : REF_TO BYTE;
// 	ptm : REF_TO BYTE;
// 	pt1, pt2 : REF_TO BYTE;
// 	su : STRING(2);
// 	pos : INT;
// END_VAR
//
// PT := REF(str);
// pto := REF(REPLACE_UML);
// ptm := pto + INT_TO_DWORD(string_length);
// pt1 := REF(su);
// pt2 := pt1 + 1;
// L := LEN(str);
// WHILE pos < L AND pos < string_length DO
// 	IF pt^ < 127 THEN
// 		(* no uml character simlply copy the character*)
// 		pto^ := pt^;
// 	ELSE
// 		(* convert the uml character *)
// 		su := TO_UML(pt^);
// 		(* we must make sure pointer are not out of range *)
// 		pto^ := pt1^;
// 		IF pto < ptm AND pt2^ > 0 THEN
// 			pto := pto + 1;
// 			pto^ := pt2^;
// 		END_IF;
// 	END_IF;
// 	(* increment pointers *)
// 	pt := pt + 1;
// 	pto := pto + 1;
// 	pos := pos + 1;
// END_WHILE;
//
// (* properly close the output string *)
// pto^ := 0;
// END_FUNCTION

FUNCTION_BLOCK TICKER

VAR_INPUT
	N : INT;
	PT : TIME;
END_VAR

VAR_IN_OUT
	Text : STRING(STRING_LENGTH);
END_VAR

VAR_OUTPUT
	Display : STRING(STRING_LENGTH);
END_VAR
VAR
	delay : TP;
	step : INT;
END_VAR

(* generate next ticker when delay is low *)
IF N < LEN(text) THEN
	IF NOT delay.Q THEN
		(* increase step for next tick *)
		step := step + 1;
		IF step > LEN(text) THEN step := 1; END_IF;
		(* extract dispay from text *)
		display := MID(text, N, step);
		(* set delay timer for next tick *)
		delay(in := TRUE, PT := PT);
	ELSE;
		(* execute delay timer *)
		delay(in := FALSE);
	END_IF;
ELSE
	display := text;
END_IF;
END_FUNCTION_BLOCK

FUNCTION TO_LOWER : BYTE
VAR_INPUT
	IN : BYTE;
END_VAR

IF in > 64 AND in < 91 THEN
   TO_LOWER := in OR 16#20;
ELSIF (in > 191 AND in < 223) AND in <> 215 AND setup.EXTENDED_ASCII THEN
   TO_LOWER := in OR 16#20;
ELSE
   TO_LOWER := in;
END_IF;
END_FUNCTION

// Commented out for beedance: it uses CHR_TO_STRING, which is commented out.
// FUNCTION TO_UML : STRING(2)
// VAR_INPUT
// 	IN : BYTE;
// END_VAR
//
// CASE in OF
// 	196:	(* Ä *)
// 		TO_UML := 'Ae';
// 	214:	(* Ö *)
// 		TO_UML := 'Oe';
// 	220:	(* Ü *)
// 		TO_UML := 'Ue';
// 	223:	(* ß *)
// 		TO_UML := 'ss';
// 	228:	(* ä *)
// 		TO_UML := 'ae';
// 	246:	(* ö *)
// 		TO_UML := 'oe';
// 	252:	(* ü *)
// 		TO_UML := 'ue';
// ELSE
// 	TO_UML := CHR_TO_STRING(IN);
// END_CASE;
// END_FUNCTION

FUNCTION TO_UPPER : BYTE
VAR_INPUT
	IN : BYTE;
END_VAR

IF in > 96 AND in < 123 THEN
   TO_UPPER := in AND 16#DF;
ELSIF in > 223 AND in <> 247 AND in <> 255 AND setup.EXTENDED_ASCII THEN
   TO_UPPER := in AND 16#DF;
ELSE
   TO_UPPER := in;
END_IF;
END_FUNCTION

FUNCTION TRIM : STRING(STRING_LENGTH)
VAR_INPUT
	str : STRING(STRING_LENGTH);
END_VAR
VAR
	pos: INT;
END_VAR

TRIM := str;
REPEAT
	pos := FIND(trim,' ');
	IF pos > 0 THEN TRIM := REPLACE(TRIM,'',1,pos); END_IF;
UNTIL pos = 0	END_REPEAT;

(* revision histroy
hm	6.10.2006		rev 1.0
	original release

hm	20. mar. 2008	rev 1.1
	avoid to call replace with pos = 0 because some systems will produce an error

hm	29. mar. 2008	rev 1.2
	changed STRING to STRING(STRING_LENGTH)
*)
END_FUNCTION

FUNCTION TRIM1 : STRING(STRING_LENGTH)
VAR_INPUT
	str : STRING(STRING_LENGTH);
END_VAR
VAR
	pos: INT;
END_VAR

TRIM1 := str;
REPEAT
	pos := FIND(trim1,'  ');
	IF pos > 0 THEN TRIM1 := REPLACE(TRIM1,' ',2,pos); END_IF;
UNTIL pos = 0	END_REPEAT;
(* beginning and ending blanks need to be stripped off *)
IF LEFT(trim1,1) = ' ' THEN trim1 := DELETE(trim1,1,1); END_IF;
IF RIGHT(trim1,1) = ' ' THEN trim1 := DELETE(trim1,1,LEN(trim1)); END_IF;

(* revision histroy
hm	4. feb. 2008    rev 1.0
	original release

hm	20. mar. 2008	rev 1.1
	avoid to call replace with pos = 0 because some systems will produce an error

hm	29. mar. 2008	rev 1.2
	changed STRING to STRING(STRING_LENGTH)
*)
END_FUNCTION

FUNCTION TRIME : STRING(string_length)
VAR_INPUT
	str : STRING(STRING_LENGTH);
END_VAR

TRIME := str;
(* beginning blanks need to be stripped off *)
WHILE LEFT(TRIME,1) = ' ' DO
	TRIME := DELETE(TRIME,1,1);
END_WHILE;

(* ending blanks need to be stripped off *)
WHILE RIGHT(TRIME,1) = ' ' DO
	TRIME := DELETE(TRIME,1,LEN(TRIME));
END_WHILE;

(* revision histroy
hm	28. mar. 2008	rev 1.0
	original release

*)
END_FUNCTION

// Commented out for beedance: it computes with pointers as addresses (pt := pt + 1); beedance references (REF_TO) have no arithmetic.
// FUNCTION UPPERCASE : STRING(STRING_LENGTH)
// VAR_INPUT
// 	str : STRING(STRING_LENGTH);
// END_VAR
// VAR
// 	pt : REF_TO BYTE;
// 	pos: INT;
// 	l: INT;
// END_VAR
//
// pt := REF(UPPERCASE);
// UPPERCASE := str;
// l := LEN(str);
// FOR pos := 1 TO l DO
// 	pt^ := TO_UPPER(pt^);
// 	pt := pt + 1;
// END_FOR;
//
// (* revision histroy
// hm	6. oct. 2006	rev 1.0
// 	original release
//
// hm	4. feb. 2008	rev 1.1
// 	improved performance
// 	added Ä,Ö,Ü
//
// hm	6. mar. 2008	rev 1.2
// 	added support for exteded Ascii
//
// hm	29. mar. 2008	rev 1.3
// 	changed STRING to STRING(STRING_LENGTH)
//
// *)
//
// END_FUNCTION

FUNCTION WEEKDAY_TO_STRING : STRING(10)
VAR_INPUT
	WDAY : INT;
	LANG : INT;
	LX : INT;
END_VAR
VAR
	ly : INT;
END_VAR

IF LANG = 0 THEN ly := LANGUAGE.DEFAULT; ELSE ly := MIN(LANG, LANGUAGE.LMAX); END_IF;
IF wday < 1 OR wday > 7 THEN
	RETURN;
ELSIF LX = 0 THEN
	WEEKDAY_TO_STRING := language.WEEKDAYS[ly, WDAY];
ELSIF Lx = 2 THEN
	WEEKDAY_TO_STRING := language.WEEKDAYS2[ly, WDAY];
END_IF;

(* revisison history

hm	21. sep. 2008	rev 1.0
	original version

hm	19. oct. 2008	rev 1.1
	changed language setup constants
*)
END_FUNCTION

FUNCTION_BLOCK CALENDAR_CALC
VAR_INPUT
	SPE : BOOL;
	H : REAL := -0.83333333333;
END_VAR
VAR_IN_OUT
	XCAL : CALENDAR;
	HOLIDAYS : ARRAY[0..29] OF HOLIDAY_DATA;
END_VAR
VAR
	last : DT;
	last_day : DINT;
	holy : HOLIDAY;
	sun : SUN_TIME;
	last_hour: INT;
	utod: TOD;
	pos : SUN_POS;
	plast: DT;
END_VAR
VAR_TEMP
	dtemp : DINT;
	tmp : INT;
END_VAR

IF xcal.UTC <> last THEN
	(* run once per second *)
	(* update utc last calculated  *)
	last := XCAL.UTC;
	utod := DT_TO_TOD(xcal.UTC);

	(* calculate ltc from utc *)
	XCAL.LOCAL_DT := UTC_TO_LTIME(XCAL.UTC, XCAL.DST_EN, XCAL.OFFSET);
	XCAL.LOCAL_DATE := DT_TO_DATE(XCAL.LOCAL_DT);
	XCAL.LOCAL_TOD := DT_TO_TOD(XCAL.LOCAL_DT);
	dtemp := DAY_OF_DATE(XCAL.LOCAL_DATE);
	xcal.night := XCAL.LOCAL_TOD < XCAL.SUN_RISE OR XCAL.LOCAL_TOD > XCAL.SUN_SET;

	(* run once per hour *)
	tmp := HOUR(xcal.LOCAL_TOD);
	IF  tmp <> last_hour THEN
		XCAL.DST_ON := DST(XCAL.UTC) AND xcal.DST_EN;
		last_hour := tmp;
	END_IF;

	(* run once per day *)
	IF dtemp <> last_day THEN
		last_day := dtemp;
		(* a new day has started, recalculate daily events *)
		XCAL.YEAR := YEAR_OF_DATE(XCAL.LOCAL_DATE);
		XCAL.MONTH := MONTH_OF_DATE(XCAL.LOCAL_DATE);
		XCAL.DAY := DAY_OF_MONTH(XCAL.LOCAL_DATE);
		XCAL.WEEKDAY := DAY_OF_WEEK(XCAL.LOCAL_DATE);
		HOLY(date_in := XCAL.LOCAL_DATE, LANGU := xcal.LANGUAGE, HOLIDAYS := HOLIDAYS);
		XCAL.HOLIDAY := HOLY.Y;
		XCAL.HOLY_NAME := HOLY.NAME;
		sun(latitude := XCAL.LATITUDE, longitude := xcal.LONGITUDE, utc := DT_TO_DATE(xcal.UTC), H := H);
		XCAL.SUN_RISE := DINT_TO_TOD(TOD_TO_DINT(sun.sun_rise) + XCAL.OFFSET * 60000 + SEL(XCAL.DST_ON,DINT#0,3600000));
		XCAL.SUN_SET := DINT_TO_TOD(TOD_TO_DINT(sun.sun_set) + XCAL.OFFSET * 60000 + SEL(XCAL.DST_ON,DINT#0,3600000));
		XCAL.SUN_MIDDAY := DINT_TO_TOD(TOD_TO_DINT(sun.MIDDAY) + XCAL.OFFSET * 60000 + SEL(XCAL.DST_ON,DINT#0,3600000));
		XCAL.SUN_HEIGTH := sun.sun_declination;
		XCAL.WORK_WEEK := WORK_WEEK(XCAL.LOCAL_DATE);
	END_IF;

	(* calculate the suns position every 10 seconds when SPE = TRUE *)
	IF SPE AND xcal.UTC -  plast >= t#25s THEN
		plast := last;
		pos(latitude := xcal.LATITUDE, longitude := xcal.LONGITUDE, utc := xcal.UTC);
		xcal.SUN_HOR := pos.B;
		xcal.SUN_VER := pos.HR;
	END_IF;
END_IF;
END_FUNCTION_BLOCK

FUNCTION DATE_ADD : DATE
VAR_INPUT
	IDATE : DATE;
	D : INT;
	W : INT;
	M : INT;
	Y : INT;
END_VAR
VAR
	mo: INT;
	yr : INT;
	dm: INT;
END_VAR

DATE_ADD := UDINT_TO_DATE(DATE_TO_UDINT(IDATE) + INT_TO_UDINT(D + W * 7) * UDINT#86400);
yr := Y + YEAR_OF_DATE(DATE_ADD);
mo := M + MONTH_OF_DATE(DATE_ADD);
dm := DAY_OF_MONTH(DATE_ADD);
WHILE mo > 12 DO
	mo := mo - 12;
	yr := yr + 1;
END_WHILE;
WHILE mo < 1 DO
	mo := mo + 12;
	yr := yr - 1;
END_WHILE;
DATE_ADD := SET_DATE(yr, mo, dm);
END_FUNCTION

FUNCTION DAY_OF_DATE : DINT
VAR_INPUT
	idate : DATE;
END_VAR

DAY_OF_DATE := UDINT_TO_DINT(DATE_TO_UDINT(idate) / 86400);
END_FUNCTION

FUNCTION DAY_OF_MONTH : INT
VAR_INPUT
	IDATE : DATE;
END_VAR
VAR
	leap: INT;
END_VAR

(* calculate the day in the year *)
DAY_OF_MONTH := DAY_OF_YEAR(idate);
(* leap will be set to one for a leap year *)
leap := BOOL_TO_INT(LEAP_OF_DATE(idate));
(* if leap year deduct one from the days of the year *)
DAY_OF_MONTH := DAY_OF_MONTH - leap;
(* search if we are in month december to march ? *)
IF DAY_OF_MONTH > setup.MTH_OFS[9] THEN
	IF DAY_OF_MONTH > setup.MTH_OFS[11] THEN
		IF DAY_OF_MONTH > setup.mth_ofs[12] THEN
			DAY_OF_MONTH := DAY_OF_MONTH - setup.MTH_OFS[12];
		ELSE
			DAY_OF_MONTH := DAY_OF_MONTH - setup.MTH_OFS[11];
		END_IF;
	ELSE
		IF DAY_OF_MONTH > setup.mth_ofs[10] THEN
			DAY_OF_MONTH := DAY_OF_MONTH - setup.MTH_OFS[10];
		ELSE
			DAY_OF_MONTH := DAY_OF_MONTH - setup.MTH_OFS[9];
		END_IF;
	END_IF;
ELSIF DAY_OF_MONTH > setup.MTH_OFS[5] THEN
	IF DAY_OF_MONTH > setup.MTH_OFS[7] THEN
		IF DAY_OF_MONTH > setup.mth_ofs[8] THEN
			DAY_OF_MONTH := DAY_OF_MONTH - setup.MTH_OFS[8];
		ELSE
			DAY_OF_MONTH := DAY_OF_MONTH - setup.MTH_OFS[7];
		END_IF;
	ELSE
		IF DAY_OF_MONTH > setup.mth_ofs[6] THEN
			DAY_OF_MONTH := DAY_OF_MONTH - setup.MTH_OFS[6];
		ELSE
			DAY_OF_MONTH := DAY_OF_MONTH - setup.MTH_OFS[5];
		END_IF;
	END_IF;
ELSIF DAY_OF_MONTH > setup.MTH_OFS[3] THEN
	IF DAY_OF_MONTH > setup.MTH_OFS[4] THEN
		DAY_OF_MONTH := DAY_OF_MONTH - setup.MTH_OFS[4];
	ELSE
		DAY_OF_MONTH := DAY_OF_MONTH - setup.MTH_OFS[3];
	END_IF;
ELSE
	(* since now we must be in february or january we need to add leap again *)
	DAY_OF_MONTH := DAY_OF_MONTH + leap;
	IF DAY_OF_MONTH > setup.MTH_OFS[2] THEN DAY_OF_MONTH := DAY_OF_MONTH - setup.mth_ofs[2]; END_IF;
	(* since nothing was true before, day_of_month must already be good *)
END_IF;

END_FUNCTION

FUNCTION DAY_OF_WEEK : INT
VAR_INPUT
	IDATE : DATE;
END_VAR

DAY_OF_WEEK := UDINT_TO_INT((DATE_TO_UDINT(idate) / 86400 + 3) MOD 7) + 1;

END_FUNCTION

FUNCTION DAY_OF_YEAR : INT
VAR_INPUT
	IDATE : DATE;
END_VAR

DAY_OF_YEAR := UDINT_TO_INT((DATE_TO_UDINT(idate) / UDINT#86400) MOD UDINT#1461);
IF DAY_OF_YEAR > 729 THEN
	IF DAY_OF_YEAR > 1095 THEN DAY_OF_YEAR := DAY_OF_YEAR - 1095; ELSE DAY_OF_YEAR := DAY_OF_YEAR - 729; END_IF;
ELSIF DAY_OF_YEAR > 364 THEN
	DAY_OF_YEAR := DAY_OF_YEAR - 364;
ELSE
	DAY_OF_YEAR := DAY_OF_YEAR + 1;
END_IF;

(*
DAY_OF_YEAR := DWORD_TO_INT((DATE_TO_DWORD(idate) - DATE_TO_DWORD(YEAR_BEGIN(YEAR_OF_DATE(idate)))) / 86400) + 1;
*)

(* revivision history
hm	4. aug. 2007		rev 1.0
	original version

hm	1. oct. 2007		rev 1.1
	added compatibility to STEP7

hm	4. jan. 2008		rev 1.2
	changed code for better performance

hm	7. oct. 2008		rev 1.3
	changed name of function year to year_of_date

hm	28. jan. 2011	rev 1.4
	improved code
*)
END_FUNCTION

FUNCTION DAY_TO_TIME : TIME
VAR_INPUT
	IN : REAL;
END_VAR

DAY_TO_TIME := DWORD_TO_TIME(REAL_TO_DWORD(IN * 86400000.0));
END_FUNCTION

FUNCTION DAYS_DELTA : DINT
VAR_INPUT
	date_1 : DATE;
	date_2 : DATE;
END_VAR

IF DATE_1 > DATE_2 THEN
	DAYS_DELTA := - UDINT_TO_DINT((DATE_TO_UDINT(date_1) - DATE_TO_UDINT(date_2)) / 86400);
ELSE
	DAYS_DELTA := UDINT_TO_DINT((DATE_TO_UDINT(date_2) - DATE_TO_UDINT(date_1)) / 86400);
END_IF;
END_FUNCTION

FUNCTION DAYS_IN_MONTH : INT
VAR_INPUT
	IDATE : DATE;
END_VAR

DAYS_IN_MONTH := DAY_OF_YEAR(IDATE);
IF LEAP_OF_DATE(IDATE) THEN
	CASE DAYS_IN_MONTH OF
		32..60	:	DAYS_IN_MONTH := 29;
		92..121 :	DAYS_IN_MONTH := 30;
		153..182:	DAYS_IN_MONTH := 30;
		245..274:	DAYS_IN_MONTH := 30;
		306..335:	DAYS_IN_MONTH := 30;
	ELSE
		DAYS_IN_MONTH := 31;
	END_CASE;
ELSE
	CASE DAYS_IN_MONTH OF
		32..59	:	DAYS_IN_MONTH := 28;
		91..120 :	DAYS_IN_MONTH := 30;
		152..181:	DAYS_IN_MONTH := 30;
		244..273:	DAYS_IN_MONTH := 30;
		305..334:	DAYS_IN_MONTH := 30;
	ELSE
		DAYS_IN_MONTH := 31;
	END_CASE;
END_IF;
END_FUNCTION

FUNCTION DAYS_IN_YEAR : INT
VAR_INPUT
	IDATE : DATE;
END_VAR

IF LEAP_OF_DATE(IDATE) THEN
	DAYS_IN_YEAR := 366;
ELSE
	DAYS_IN_YEAR := 365;
END_IF;
END_FUNCTION

FUNCTION_BLOCK DCF77
VAR_INPUT
	REC : BOOL;
	SET : BOOL;
	SDT : DT;
	DSI : BOOL;
END_VAR
VAR_INPUT CONSTANT
	SYNC_TIMEOUT : TIME := t#2m;
	TIME_OFFSET : INT := 1;
	DST_EN : BOOL := TRUE;
END_VAR
VAR_OUTPUT
	TP : BOOL;
	DS : BOOL;
	WDAY : INT;
	ERROR : BOOL := TRUE;
	RTC : DT;
	RTC1 : DT;
	MSEC : INT;
	SYNC : BOOL;
END_VAR
VAR
	mez : DT;
	utc : DT;
	state : INT;
	edge: BOOL;
	tx : TIME;
	ty: TIME;
	last : TIME;
	bits : ARRAY[0..58] OF BOOL;
	cnt : INT;
	i : INT;
	old_time : DT;
	minute : INT;
	hour : INT;
	day : INT;
	month : INT;
	year : INT;
	last_sync: TIME;
	t1: TIME;
	tz: TIME;
	init: BOOL;
END_VAR

(* if tp was set it should only be active for 1 cycle *)
TP := FALSE;

(* read system time *)
t1 := DWORD_TO_TIME(T_PLC_MS());
tx := t1 - last;

IF rec XOR edge THEN
	edge := rec;
	IF NOT rec AND tx > t#1700ms AND tx < t#2000ms THEN
		(* start condition reached *)
		state := 0;
		tp := NOT error;
	ELSIF NOT rec AND tx > t#700ms AND tx < t#1000ms THEN
		(* second switch detected *)
		IF state < 58 THEN state := state +1; ELSE state := 0; END_IF;
	ELSIF rec AND tx  < t#120ms THEN
		(* bit 0 detected  *)
		bits[state] := 0;
	ELSIF rec AND tx > t#120ms AND tx < t#250ms THEN
		(* bit 1 detected *)
		bits[state] := 1;
	ELSE
		(* error condition received signal is not valid *)
		error := TRUE;
		state := 0;
	END_IF;
	last := last + tx;
	IF rec AND state = 58 THEN
		error := FALSE;

		(* decode the bits and check for possible errors *)
		IF bits[0] OR NOT (bits[17] XOR bits[18]) OR NOT bits[20] THEN error := TRUE; END_IF;
		(* decode minute *)
		MINUTE := 0;
		MINUTE.0 := bits[21];
		MINUTE.1 := bits[22];
		MINUTE.2 := bits[23];
		MINUTE.3 := bits[24];
		IF bits[25] THEN MINUTE := MINUTE + 10; END_IF;
		IF bits[26] THEN MINUTE := MINUTE + 20; END_IF;
		IF bits[27] THEN MINUTE := MINUTE + 40; END_IF;
		IF MINUTE > 59 OR (bits[21] XOR bits[22] XOR bits[23] XOR bits[24] XOR bits[25] XOR bits[26] XOR bits[27] XOR bits[28]) THEN error := TRUE; END_IF;

		(* decode hour *)
		HOUR := 0;
		HOUR.0 := bits[29];
		HOUR.1 := bits[30];
		HOUR.2 := bits[31];
		HOUR.3 := bits[32];
		IF bits[33] THEN HOUR := HOUR + 10; END_IF;
		IF bits[34] THEN HOUR := HOUR +20; END_IF;
		IF HOUR > 23 OR (bits[29] XOR bits[30] XOR bits[31] XOR bits[32] XOR bits[33] XOR bits[34] XOR bits[35]) THEN error := TRUE; END_IF;

		(* decode day of month *)
		day := 0;
		day.0 := bits[36];
		day.1 := bits[37];
		day.2 := bits[38];
		day.3 := bits[39];
		IF bits[40] THEN day := day + 10; END_IF;
		IF bits[41] THEN day := day + 20; END_IF;
		IF day > 31 THEN error := TRUE; END_IF;

		(* decode day of week *)
		wday := 0;
		wday.0 := bits[42];
		wday.1 := bits[43];
		wday.2 := bits[44];
		IF wday > 7 OR wday < 1 THEN error := TRUE; END_IF;

		(* decode month *)
		MONTH := 0;
		MONTH.0 := bits[45];
		MONTH.1 := bits[46];
		MONTH.2 := bits[47];
		MONTH.3 := bits[48];
		IF bits[49] THEN MONTH := MONTH +10; END_IF;
		IF MONTH > 12 THEN error := TRUE; END_IF;

		(* decode year *)
		YEAR := 0;
		YEAR.0 := bits[50];
		YEAR.1 := bits[51];
		YEAR.2 := bits[52];
		YEAR.3 := bits[53];
		IF bits[54] THEN YEAR := YEAR + 10; END_IF;
		IF bits[55] THEN YEAR := YEAR + 20; END_IF;
		IF bits[56] THEN YEAR := YEAR + 40; END_IF;
		IF bits[57] THEN YEAR := YEAR + 80; END_IF;

		(* check parity for bits 36 to 58 *)
		cnt := 0;
		FOR i := 36 TO 58 DO IF bits[i] THEN cnt := cnt + 1; END_IF; END_FOR;
		IF NOT EVEN(cnt) THEN error := TRUE; END_IF;

		(* time must be valid for two cycles to clear error flag *)
		IF NOT error THEN
			(* set outputs *)
			old_time := mez;
			IF YEAR >= 70 THEN YEAR := YEAR + 1900; ELSE YEAR := YEAR + 2000; END_IF;
			mez := SET_DT(YEAR,MONTH,day,HOUR,MINUTE,0);
			DS := bits[17];
			IF DS THEN
				UTC := UDINT_TO_DT(DT_TO_UDINT(mez) - 7200);
			ELSE
				UTC := UDINT_TO_DT(DT_TO_UDINT(mez) - 3600);
			END_IF;

			(* set trigger signal only if the receiver has received 2 successive minutes *)
			IF mez <> old_time + t#1m THEN error := TRUE ; END_IF;
		END_IF;
	END_IF;
END_IF;

(* this portion implements a free running clock which is triggered by the dcf77 signal *)
tz := UDINT_TO_TIME(INT_TO_UDINT(ABS(time_offset)) * 3600000);

(* input sdt is copied to utc at first power up *)
IF NOT init OR SET THEN
	init := TRUE;
	utc := sdt;
	tp := TRUE;
	DS := DSI;
END_IF;

IF tp THEN
	rtc := utc;
	IF DS AND dst_en THEN
		IF time_offset < 0 THEN	rtc1 := rtc - tz + t#1h; ELSE rtc1 := rtc + tz + t#1h; END_IF;
	ELSE
		IF time_offset < 0 THEN rtc1 := rtc - tz; ELSE rtc1 := rtc + tz; END_IF;
	END_IF;
	sync := TRUE;
	last_sync := last;
	ty := last;
ELSIF rtc > DWORD_TO_DT(0) AND T1 - ty >= t#1s THEN
	rtc := rtc + t#1s;
	rtc1 := rtc1 + t#1s;
	ty := ty + t#1s;
	sync := ty - last_sync < sync_timeout AND last_sync > DWORD_TO_TIME(0);
	wday := DAY_OF_WEEK(DT_TO_DATE(rtc1));
	DS := dst_en AND DST(utc);
END_IF;
msec := TIME_TO_INT(t1 - ty);

(* decode information
bits		content
0			Bitwert immer 0
1 bis 14	reserviert für Betriebsinformationen (nicht für DCF77-Nutzer bestimmt)
15			Rufbit für Alarmierung der PTB-Mitarbeiter
			(bis Mai 2003: Bitwert = 0 falls normale Antenne in Verwendung; 1 = Backupantenne)
16			Bitwert = 1 falls ein Wechsel von MEZ nach MESZ oder umgekehrt bevorsteht; Dauer der Anzeige: 1 Stunde
17 + 18	gültige Zeit = MEZ, falls Bit 17=0 und Bit 18=1
			gültige Zeit = MESZ, falls Bit 17=1 und Bit 18=0
19			Bitwert = 1 falls innerhalb den nächsten 59 Minuten eine Schaltsekunde angeordnet ist. Beim Einfügen einer Schaltsekunde wird anstelle der 59. die 60. Sekundenmarke weggelassen und in der 58. erfolgt ausnahmsweise ein Trägerabfall.
20			Startbit für Zeitinformation (immer 1)
21 - 27		1, 2, 4, 8, 10, 20, 40 Minuten (bitweise Addition)
28			Prüfbit (gerade Parität) für die Bits 21-27
29 - 34		1, 2, 4, 8, 10, 20 Stunden (bitweise Addition)
35			Prüfbit (gerade Parität) für die Bits 29-34
36 - 41		Tagesnummer im aktuellen Monat: 1, 2, 4, 8, 10, 20 (bitweise Addition)
42 - 44		Tagesnummer in der aktuellen Woche: 1, 2, 4 (bitweise Addition)
45 - 49		Monatsnummer: 1, 2, 4, 8, 10 (bitweise Addition)
50 - 57		Jahr (zweistellig): 1, 2, 4, 8, 10, 20, 40, 80 (bitweise Addition)
58			Prüfbit (gerade Parität) füR die Bits 36-57

*)

END_FUNCTION_BLOCK

FUNCTION DST : BOOL
VAR_INPUT
	UTC : DT;
END_VAR
VAR
	yr : INT;
	yr4 : DWORD;
	ltc: DWORD;
	idate : DWORD;
END_VAR
